(* Logix 5000 project; controller CIP vendor 1 type 14 code 106 rev 20.12; software revision 20.06 *)

TASK MainTask (continuous, watchdog 500 ms) : MainProgram

MODULES
   Local : vendor 1 type 14 code 106 (Compact 0, rev 20.12)
      Digital_Input_2 : 1769-IQ16 (Compact 5, rev 3.1, Input RPI 20 ms)
      Digital_Input_3 : 1769-IQ16 (Compact 6, rev 3.1, Input RPI 20 ms)
      Digital_Input_1 : 1769-IQ16 (Compact 4, rev 3.1, Input RPI 20 ms)
      Analog_Output_1 : vendor 1 type 10 code 45 (Compact 3, rev 2.1, Output RPI 80 ms)
      Analog_Input_1 : 1769-IF8 (Compact 1, rev 1.1, Output RPI 80 ms)
      Digital_Output_2 : 1769-OB16 (Compact 8, rev 3.1, Output RPI 20 ms)
      Analog_Input_2 : 1769-IF8 (Compact 2, rev 1.1, Output RPI 80 ms)
      Digital_Output_1 : 1769-OB16 (Compact 7, rev 3.1, Output RPI 20 ms)
      WASHER : 1734-AENT (Ethernet 192.168.1.58, rev 4.3, Output RPI 20 ms)
         Washer_Digital_Input_3 : 1734-IB8 (PointIO 5, rev 3.22)
         Washer_Digital_Input_1 : 1734-IB8 (PointIO 3, rev 3.22)
         Washer_Digital_Input_2 : 1734-IB8 (PointIO 4, rev 3.22)
         Washer_Analog_Input_1 : vendor 1 type 115 code 210 (PointIO 1, rev 3.2, Input RPI 80 ms)
         Washer_Digital_Output_2 : 1734-OB8 (PointIO 7, rev 3.22)
         Washer_Analog_Output_1 : 1734-OE2C (PointIO 2, rev 3.5, Output RPI 80 ms)
         Washer_Digital_Output_3 : 1734-OB8 (PointIO 8, rev 3.22)
         Washer_Digital_Output_1 : 1734-OB8 (PointIO 6, rev 3.22)
END_MODULES

TYPE Produce_Consume_Data :
STRUCT
   CommStatus : CONNECTION_STATUS;
   String : STRING[2];
   Real : REAL[10];
   DINT : DINT[10];
END_STRUCT
END_TYPE

TYPE RECIPE :
STRUCT
   OpCode : DINT[97];
   StepTime : DINT[97];
   Setpoint : REAL[97];
   Name : STRING;
END_STRUCT
END_TYPE

TYPE Security_Main_HMI :
STRUCT
   Timers : TIMER[10];
   Bits : DINT;
   Counters : COUNTER[6];
   User_Security_Name : STRING;
   User_Security_Name_Display : STRING[2];
   User_Security_Name_Temp : STRING;
   User_Security_Password : STRING;
   User_Security_Password_Temp : STRING;
   User_Security_Level : DINT;
   Number_Of_Users : DINT;
   User_Names : STRING[53];
   User_Names_Edit : STRING[53];
   User_Passwords : STRING[53];
   User_Passwords_Edit : STRING[53];
   User_Security_Levels : DINT[53];
   User_Security_Levels_Edit : DINT[53];
   Security_Save_Edit_Changes : BOOL;
   Security_Login_Enter_User_Button : BOOL;
   Security_Logout_Button : BOOL;
   Control_1 : CONTROL;
   Control_2 : CONTROL;
   Control_3 : CONTROL;
   User_Security_Name_Clear : STRING;
   User_Security_Password_Clear : STRING;
   Security_Login_Enter_Password_Button : BOOL;
   Name_Temp : DINT;
   Password_Temp : DINT;
   Auto_Logout_Counter : COUNTER;
   Auto_Logout_Timer_Enable : BOOL;
   Auto_Logout_Timer_Enabled : BOOL;
   Auto_Logout_Preset : DINT;
   Auto_Logout_Temp : DINT;
   PanelView_Control : DINT;
   PanelView_Status : DINT;
   PanelView_Security_Edit_Active : BOOL;
   PanelView_Security_Password_Length : DINT;
END_STRUCT
END_TYPE

TYPE Security_Remote_HMI :
STRUCT
   Timers : TIMER[3];
   Bits : DINT;
   User_Security_Name : STRING;
   User_Security_Name_Display : STRING[2];
   User_Security_Name_Temp : STRING;
   User_Security_Password : STRING;
   User_Security_Password_Temp : STRING;
   User_Security_Level : DINT;
   Number_Of_Users : DINT;
   User_Names : STRING[53];
   User_Passwords : STRING[53];
   User_Security_Levels : DINT[53];
   Security_Login_Enter_User_Button : BOOL;
   Security_Logout_Button : BOOL;
   Control_1 : CONTROL;
   User_Security_Name_Clear : STRING;
   User_Security_Password_Clear : STRING;
   Security_Login_Enter_Password_Button : BOOL;
   Auto_Logout_Counter : COUNTER;
   Auto_Logout_Timer_Enable : BOOL;
   Auto_Logout_Timer_Enabled : BOOL;
   Auto_Logout_Temp : DINT;
   PanelView_Control : DINT;
   PanelView_Status : DINT;
END_STRUCT
END_TYPE

VAR_GLOBAL   (* controller tags *)
   Alarm_Ack : INT[8];
   Alarm_Ack_All_PB : BOOL;
   Alarm_Present : INT[8] := ([0] := 70, [7] := 16384);
   Alarm_Preset_Indx : DINT := 118;
   Alarm_Remote_Ack_All : BOOL;
   Alarm_Status_Reset : BOOL;
   Alarm_Timer : TIMER[128] := ([0].PRE := 1500, [1].ACC := 4, [1].EN := 1, [1].DN := 1, [2].ACC := 4, [2].EN := 1, [2].DN := 1, [6].PRE := 3000, [7].PRE := 5000, [8].PRE := 5000, [9].PRE := 5000, [10].PRE := 5000, [11].PRE := 5000, [12].PRE := 5000, [13].PRE := 5000, [14].PRE := 5000, [15].PRE := 5000, [16].PRE := 5000, [17].PRE := 5000, [17].ACC := 5000, [17].EN := 1, [17].DN := 1, [18].PRE := 3000000, [19].PRE := 300000, [20].PRE := 1000, [21].PRE := 5000, [22].PRE := 1000, [23].PRE := 300000, [24].PRE := 900000, [25].PRE := 900000, [26].PRE := 300000, [27].PRE := 300000, [28].PRE := 500, [29].PRE := 500, [30].PRE := 8000, [31].PRE := 15000, [32].PRE := 8000, [33].PRE := 15000, [34].PRE := 8000, [35].PRE := 15000, [36].PRE := 8000, [37].PRE := 15000, [38].PRE := 5000, [39].PRE := 5000, [40].PRE := 3000, [41].PRE := 3000, [42].PRE := 3000, [44].PRE := 300000, [45].PRE := 5000, [45].ACC := 5001, [45].EN := 1, [45].DN := 1, [46].PRE := 8000, [47].PRE := 15000, [48].PRE := 8000, [49].PRE := 15000, [50].PRE := 5000, [51].PRE := 5000, [52].PRE := 5000, [53].PRE := 5000,
        [54].PRE := 5000, [55].PRE := 5000, [56].PRE := 5000, [57].PRE := 5000, [58].PRE := 5000, [59].PRE := 5000, [60].PRE := 5000, [61].PRE := 5000, [62].PRE := 5000, [63].PRE := 5000, [64].PRE := 5000, [65].PRE := 5000, [66].PRE := 5000, [67].PRE := 5000, [68].PRE := 5000, [69].PRE := 5000, [70].PRE := 5000, [71].PRE := 5000, [72].PRE := 5000, [73].PRE := 5000, [74].PRE := 5000, [75].PRE := 5000, [76].PRE := 5000, [77].PRE := 5000, [78].PRE := 5000, [78].ACC := 5001, [78].EN := 1, [78].DN := 1, [79].PRE := 5000, [79].ACC := 5001, [79].EN := 1, [79].DN := 1, [80].PRE := 5000, [81].PRE := 5000, [82].PRE := 5000, [83].PRE := 5000, [83].ACC := 5001, [83].EN := 1, [83].DN := 1, [84].PRE := 3000, [85].PRE := 3000, [85].ACC := 3002, [85].EN := 1, [85].DN := 1, [86].PRE := 1000, [87].PRE := 3000, [88].PRE := 10000, [89].PRE := 1800000, [90].PRE := 3000, [91].PRE := 3000, [93].PRE := 20000, [94].PRE := 10000, [95].PRE := 1000, [96].PRE := 5000, [96].ACC := 5001, [96].EN := 1, [96].DN := 1, [97].PRE := 5000, [97].ACC := 5001, [97].EN := 1,
        [97].DN := 1, [98].PRE := 5000, [98].ACC := 5001, [98].EN := 1, [98].DN := 1, [99].PRE := 5000, [99].ACC := 5001, [99].EN := 1, [99].DN := 1, [100].PRE := 10000, [101].PRE := 10000, [102].PRE := 10000, [103].PRE := 10000, [104].PRE := 5000, [105].PRE := 5000, [106].PRE := 5000, [107].PRE := 5000, [108].PRE := 5000, [109].PRE := 5000, [110].PRE := 5000, [111].PRE := 5000, [112].PRE := 5000, [113].PRE := 5000, [114].PRE := 5000, [114].ACC := 5001, [114].EN := 1, [114].DN := 1, [115].PRE := 5000, [115].ACC := 5001, [115].EN := 1, [115].DN := 1, [116].PRE := 8000, [117].PRE := 15000, [118].PRE := 8000, [119].PRE := 15000, [120].PRE := 8000, [121].PRE := 15000, [122].PRE := 8000, [123].PRE := 15000, [124].PRE := 5000, [124].ACC := 5001, [124].EN := 1, [124].DN := 1, [125].PRE := 5000, [125].ACC := 5001, [125].EN := 1, [125].DN := 1, [126].PRE := 5000, [126].ACC := 576, [126].EN := 1, [126].TT := 1, [127].PRE := 5000, [127].ACC := 5001, [127].EN := 1, [127].DN := 1);
   Alarm_Timer_Preset : DINT[128] := ([6] := 3000, [7] := 5000, [8] := 5000, [9] := 5000, [10] := 5000, [11] := 5000, [12] := 5000, [13] := 5000, [14] := 5000, [15] := 5000, [16] := 5000, [17] := 5000, [18] := 3000000, [19] := 300000, [20] := 1000, [21] := 5000, [22] := 1000, [23] := 300000, [24] := 900000, [25] := 900000, [26] := 300000, [27] := 300000, [28] := 500, [29] := 500, [30] := 8000, [31] := 15000, [32] := 8000, [33] := 15000, [34] := 8000, [35] := 15000, [36] := 8000, [37] := 15000, [38] := 5000, [39] := 5000, [40] := 3000, [41] := 3000, [42] := 3000, [44] := 300000, [45] := 5000, [46] := 8000, [47] := 15000, [48] := 8000, [49] := 15000, [50] := 5000, [51] := 5000, [52] := 5000, [53] := 5000, [54] := 5000, [55] := 5000, [56] := 5000, [57] := 5000, [58] := 5000, [59] := 5000, [60] := 5000, [61] := 5000, [62] := 5000, [63] := 5000, [64] := 5000, [65] := 5000, [66] := 5000,
        [67] := 5000, [68] := 5000, [69] := 5000, [70] := 5000, [71] := 5000, [72] := 5000, [73] := 5000, [74] := 5000, [75] := 5000, [76] := 5000, [77] := 5000, [78] := 5000, [79] := 5000, [80] := 5000, [81] := 5000, [82] := 5000, [83] := 5000, [84] := 3000, [85] := 3000, [86] := 1000, [87] := 3000, [88] := 10000, [89] := 1800000, [90] := 3000, [91] := 3000, [93] := 20000, [94] := 10000, [95] := 1000, [96] := 5000, [97] := 5000, [98] := 5000, [99] := 5000, [100] := 10000, [101] := 10000, [102] := 10000, [103] := 10000, [104] := 5000, [105] := 5000, [106] := 5000, [107] := 5000, [108] := 5000, [109] := 5000, [110] := 5000, [111] := 5000, [112] := 5000, [113] := 5000, [114] := 5000, [115] := 5000, [116] := 8000, [117] := 15000, [118] := 8000, [119] := 15000, [120] := 8000, [121] := 15000, [122] := 8000, [123] := 15000, [124] := 5000, [125] := 5000, [126] := 5000, [127] := 5000);
   Bit : BOOL[128] := ([10] := 1, [15] := 1, [16] := 1, [30] := 1, [34] := 1, [35] := 1, [37] := 1, [40] := 1, [41] := 1, [49] := 1, [52] := 1, [54] := 1, [55] := 1, [60] := 1, [66] := 1, [68] := 1, [70] := 1, [81] := 1, [82] := 1, [100] := 1);
   Counter : COUNTER[10] := ([1].PRE := 9999, [1].ACC := 1, [2].PRE := 4, [3].PRE := 3, [5].PRE := 64, [5].ACC := 12, [6].PRE := 20);
   IN_F8_50_99 : REAL[50] := ([0] := nan); {produced}
   IN_N7_100_199 : INT[100] := ([0] := 35, [1] := 1, [50] := 22428, [51] := -3734, [52] := 32, [53] := -32768, [54] := 12, [55] := -32768, [56] := 11180, [57] := -3792, [58] := 4804, [59] := 976, [60] := 16578, [61] := 20792, [62] := 1, [64] := 4, [66] := 3, [74] := 1, [76] := 12, [77] := -32768, [78] := 12, [79] := -32768, [80] := 11180, [81] := -3792, [82] := 30396, [83] := 1, [84] := 16578, [85] := 19059, [86] := 1, [88] := 4, [90] := 3); {produced}
   Integer : DINT[150] := ([0] := 1, [1] := 1, [5] := 2, [6] := 2, [7] := 1, [8] := 7, [10] := 36, [11] := 29, [12] := 65, [15] := -33, [20] := 20, [21] := 21, [22] := 61, [26] := 120, [27] := 120, [28] := 100, [29] := 1, [36] := -4, [38] := -1, [39] := 190, [40] := 80, [41] := 80, [43] := 120, [44] := 120, [45] := 120, [46] := 120, [48] := 50, [52] := 2, [53] := -2, [54] := 2, [56] := 6242, [57] := 31208, [58] := 12, [60] := 16383, [61] := 84, [62] := 10000, [80] := 5921);
   Integer_1 : ALIAS FOR Integer[1];
   Integer_6 : ALIAS FOR Integer[6];
   IO_Status : INT := 16384;
   IO_Status_Masked : INT := 16384;
   Level_Bits : BOOL[32] := ([1] := 1, [3] := 1, [4] := 1, [5] := 1, [7] := 1, [10] := 1, [11] := 1, [15] := 1, [17] := 1, [18] := 1, [19] := 1, [20] := 1);
   Level_Timers : TIMER[20] := ([0].PRE := 30000, [1].PRE := 60000, [2].PRE := 45000, [3].PRE := 75000, [3].ACC := 3, [3].EN := 1, [3].DN := 1, [4].PRE := 900000, [4].ACC := 900004, [4].EN := 1, [4].DN := 1, [5].PRE := 75000, [5].ACC := 75001, [5].EN := 1, [5].DN := 1, [7].PRE := 3000, [7].ACC := 3002, [7].EN := 1, [7].DN := 1, [8].PRE := 3000, [8].ACC := 3000, [8].EN := 1, [8].DN := 1, [10].PRE := 2000, [11].PRE := 1000, [11].ACC := 1000, [12].PRE := 1000, [12].ACC := 1000, [13].PRE := 1000, [13].ACC := 1000, [14].PRE := 1000, [14].ACC := 1000);
   Message_Index : ALIAS FOR Integer[30];
   Message_Present : INT[4] := ([1] := -32768, [3] := 2048);
   Message_SEQ : DINT[101] := ([1] := 32, [2] := 32, [3] := 14, [4] := 31, [5] := 32, [6] := 25, [7] := 36);
   Message_Timer : TIMER[1] := ([0].PRE := 1500, [0].ACC := 89, [0].EN := 1, [0].TT := 1);
   Minor_Faults : DINT;
   MOA_OFF : DINT[10] := ([1] := 2112);
   MOA_ON : DINT[10] := ([1] := 8320, [2] := 1536);
   MOA_ONS : DINT;
   MOA_Screen1_Auto : BOOL;
   MOA_Screen1_Man_Off : BOOL;
   MOA_Screen1_Man_On : BOOL;
   MOA_Screen2_Auto : BOOL;
   MOA_Screen2_Man_Off : BOOL;
   MOA_Screen2_Man_On : BOOL;
   MOA_Screen3_Auto : BOOL;
   MOA_Screen3_Man_Off : BOOL;
   MOA_Screen3_Man_On : BOOL;
   MOA_Screen4_Auto : BOOL;
   MOA_Screen4_Man_Off : BOOL;
   MOA_Screen4_Man_On : BOOL;
   MOA_Select : DINT[10] := ([1] := 8192, [2] := 1024, [3] := 64, [4] := 128, [5] := 128, [6] := 1);
   MOA_SP_Supply_Pump_Speed : DINT := 35;
   MOA_Status : DINT[10] := ([1] := 10432, [2] := 1536);
   MOA_Temp : DINT := -1025;
   One_Shot : BOOL[128] := ([11] := 1, [12] := 1, [13] := 1, [14] := 1, [15] := 1, [16] := 1, [17] := 1, [29] := 1, [30] := 1, [31] := 1, [32] := 1, [50] := 1);
   OpCode_Pin : DINT[5];
   OpCode_Word : DINT[5,97] := ([1,2] := 16#0000_821c, [1,3] := 16#0000_823c, [1,4] := 16#0000_823c, [1,5] := 16#0000_2001, [1,6] := 16#0000_0004, [1,8] := 16#0000_803d, [1,9] := 16#0000_0125, [1,10] := 16#0000_0125, [1,11] := 16#0000_0125, [1,12] := 16#0000_0125, [1,13] := 16#0000_180c, [1,14] := 16#0000_180c, [1,15] := 16#0000_180c, [1,16] := 16#0000_180c, [1,17] := 16#0000_180c, [1,18] := 16#0000_180c, [1,19] := 16#0000_180c, [1,20] := 16#0000_180c, [1,21] := 16#0000_0025, [1,22] := 16#0000_0025, [1,23] := 16#0000_0025, [1,24] := 16#0000_0025, [1,25] := 16#0000_100c, [1,26] := 16#0000_100c, [1,27] := 16#0000_100c, [1,28] := 16#0000_100c, [1,29] := 16#0000_0525, [1,30] := 16#0000_0525, [1,31] := 16#0000_0525, [1,32] := 16#0000_0525, [1,33] := 16#0000_1804, [1,34] := 16#0000_1804, [1,37] := 16#0000_8224, [1,38] := 16#0000_8224, [1,39] := 16#0000_8224, [1,40] := 16#0000_8020, [1,41] := 16#0000_8020, [1,42] := 16#0000_8020, [1,43] := 16#0000_80a0, [1,44] := 16#0000_80a0, [1,45] := 16#0000_80a0, [1,46] := 16#0000_8080, [1,47] := 16#0000_8080, [1,55] := 16#0000_0005, [1,56] := 16#0000_8204, [1,57] := 16#0000_8204, [1,58] := 16#0000_0005, [1,59] := 16#0000_0005, [1,60] := 16#0000_8080, [2,6] := 16#0000_8000, [2,9] := 16#0000_c800, [2,10] := 16#0000_c800, [2,11] := 16#0000_c800, [2,12] := 16#0000_c800, [2,13] := 16#0000_c202, [2,14] := 16#0000_c202, [2,15] := 16#0000_c202, [2,16] := 16#0000_c202, [2,17] := 16#0000_c101, [2,18] := 16#0000_c101,
        [2,19] := 16#0000_c101, [2,20] := 16#0000_c101, [2,21] := 16#0000_c400, [2,22] := 16#0000_c400, [2,23] := 16#0000_c400, [2,24] := 16#0000_c400, [2,25] := 16#0000_c400, [2,26] := 16#0000_c400, [2,27] := 16#0000_c400, [2,28] := 16#0000_c400, [2,29] := 16#0000_c080, [2,30] := 16#0000_c080, [2,31] := 16#0000_c080, [2,32] := 16#0000_c080, [2,33] := 16#0000_8202, [2,34] := 16#0000_8101, [2,37] := 16#0000_c000, [2,38] := 16#0000_c000, [2,39] := 16#0000_c000, [2,40] := 16#0000_4000, [2,41] := 16#0000_4000, [2,42] := 16#0000_4000, [2,43] := 16#0000_4000, [2,44] := 16#0000_4000, [2,45] := 16#0000_4000, [2,55] := 16#0000_8800, [2,56] := 16#0000_8200, [2,57] := 16#0000_8100, [2,58] := 16#0000_8400, [2,59] := 16#0000_8080, [3,2] := 16#0000_4020, [3,3] := 16#0000_f2f0, [3,4] := 16#0000_cd30, [3,5] := 16#0000_4000, [3,6] := 16#0000_4000, [3,8] := 16#0000_0020, [3,9] := 16#0000_a200, [3,10] := 16#0000_9200, [3,11] := 16#0000_8900, [3,12] := 16#0000_8500, [3,13] := 16#0000_a200, [3,14] := 16#0000_9200, [3,15] := 16#0000_8900, [3,16] := 16#0000_8500, [3,17] := 16#0000_a200, [3,18] := 16#0000_9200, [3,19] := 16#0000_8900, [3,20] := 16#0000_8500, [3,21] := 16#0000_a200, [3,22] := 16#0000_9200, [3,23] := 16#0000_8900, [3,24] := 16#0000_8500, [3,25] := 16#0000_a200, [3,26] := 16#0000_9200, [3,27] := 16#0000_8900, [3,28] := 16#0000_8500, [3,29] := 16#0000_a200, [3,30] := 16#0000_9200, [3,31] := 16#0000_8900, [3,32] := 16#0000_8500,
        [3,33] := 16#0000_4000, [3,34] := 16#0000_4000, [3,35] := 16#0000_3210, [3,36] := 16#0000_3210, [3,37] := 16#0000_b200, [3,38] := 16#0000_8900, [3,39] := 16#0000_8500, [3,40] := 16#0000_0200, [3,41] := 16#0000_0100, [3,42] := 16#0000_0100, [3,43] := 16#0000_3200, [3,44] := 16#0000_0900, [3,45] := 16#0000_0500, [3,46] := 16#0000_2080, [3,47] := 16#0000_1040, [3,55] := 16#0000_8008, [3,56] := 16#0000_8008, [3,57] := 16#0000_8008, [3,58] := 16#0000_8008, [3,59] := 16#0000_8008, [3,60] := 16#0000_0008, [3,65] := 16#0000_0001, [3,66] := 16#0000_0001, [3,67] := 16#0000_0001, [3,68] := 16#0000_0001, [3,69] := 16#0000_0001, [4,35] := 16#0000_0003, [4,36] := 16#0000_0001, [4,49] := 16#0000_2000, [4,50] := 16#0000_1000, [4,51] := 16#0000_0800, [4,52] := 16#0000_0400, [4,53] := 16#0000_0200, [4,54] := 16#0000_0100);
   OUT_F8_0_49 : REAL[50] := ([1] := 21.79088, [2] := 22.761398, [5] := 14.0, [6] := 3.1312947, [7] := -0.5218824, [8] := -1.4997253, [9] := 0.003662333, [11] := 20.120556, [12] := 20.04044, [20] := 50.0, [30] := 60.0, [31] := 0.2, [32] := 0.1, [33] := 110.0, [34] := 195.0, [35] := 10.0, [36] := 150.0, [37] := 190.0, [38] := 60.0, [39] := 60.0, [40] := 80.0, [41] := 190.0, [42] := 5.5, [43] := 10.5); {produced}
   OUT_N7_0_99 : INT[100] := ([0] := 4, [1] := 8, [2] := 1, [6] := 32, [10] := 12, [11] := -21846, [12] := 2730, [13] := 8320, [14] := 1536, [20] := 20482, [21] := 170, [22] := 8, [30] := 70, [37] := 16384, [41] := -32768); {produced}
   Panelview : INT[40] := ([0] := 6144, [3] := 65, [8] := 1, [14] := 1, [15] := 1, [20] := 2, [31] := 1, [32] := 1, [33] := 1, [34] := -1);
   PID1 : PID := (CTL := -2080340864, EN := 1, SWM := 1, INI := 1, DVNA := 1, PVHA := 1, KP := 1.2, KI := 0.1, BIAS := 46.65812, MAXS := 100.0, MAXO := 51.0, UPD := 0.01, PV := 21.79088, ERR := -21.79088, MAXI := 100.0, MAXCV := 16383.0, MAXTIE := 16383.0, DATA[0] := -20.509062, DATA[1] := -348.65408, DATA[2] := 21.79088, DATA[3] := -21.79088, DATA[5] := 1.0, DATA[6] := 1.0, DATA[7] := 0.16, DATA[8] := 1.2, DATA[9] := 0.1, DATA[11] := 1.2, DATA[12] := 0.1, DATA[15] := 163.83, DATA[16] := 0.006103888);
   PID2 : PID := (CTL := -2080340864, EN := 1, SWM := 1, INI := 1, DVNA := 1, PVHA := 1, KP := 0.5, KI := 0.125, BIAS := 1.0468168, MAXS := 150.0, MAXO := 100.0, UPD := 0.01, PV := 3.1312947, ERR := -3.1312947, MAXI := 150.0, MAXCV := 16383.0, MAXTIE := 16383.0, DATA[0] := -0.003051877, DATA[1] := -33.40048, DATA[2] := 3.1312947, DATA[3] := -3.1312947, DATA[5] := 0.6666667, DATA[6] := 1.0, DATA[7] := 0.16, DATA[8] := 0.5, DATA[9] := 0.125, DATA[11] := 0.5, DATA[12] := 0.125, DATA[15] := 163.83, DATA[16] := 0.006103888);
   PID3 : PID := (CTL := -2080340864, EN := 1, SWM := 1, INI := 1, DVNA := 1, PVHA := 1, KP := 8.0, KI := 0.1, BIAS := 75.446365, MAXS := 150.0, DB := 3.0, MAXO := 100.0, UPD := 0.01, PV := 20.120556, ERR := -20.120556, MAXI := 150.0, MAXCV := 16383.0, MAXTIE := 16383.0, DATA[0] := 31.863266, DATA[1] := -214.61926, DATA[2] := 20.120556, DATA[3] := -20.120556, DATA[5] := 0.6666667, DATA[6] := 1.0, DATA[7] := 0.16, DATA[8] := 8.0, DATA[9] := 0.1, DATA[11] := 8.0, DATA[12] := 0.1, DATA[15] := 163.83, DATA[16] := 0.006103888);
   PID3_Timer : TIMER[4] := ([0].PRE := 5000);
   PID_Button : DINT[5];
   PID_Button_ONS : DINT[5];
   PID_ONS : DINT[5] := ([1] := 2, [2] := 10, [3] := 2, [4] := 4);
   PID_Timer : TIMER[5] := ([0].PRE := 5000, [0].ACC := 5000, [0].EN := 1, [0].DN := 1, [1].PRE := 10000, [2].PRE := 5000, [2].EN := 1, [2].DN := 1, [3].PRE := 4000, [4].PRE := 50, [4].ACC := 53, [4].EN := 1, [4].DN := 1);
   PV_Current_Select_Step_Op : DINT := 52;
   PV_Edit_Opcodes : DINT[300] := ([1] := 50, [2] := 5, [3] := 52, [4] := 12, [5] := 11, [6] := 65, [7] := 41, [8] := 5, [9] := 33, [10] := 16, [11] := 15, [12] := 67, [13] := 38, [14] := 41, [15] := 2, [16] := 8, [17] := 51, [18] := 5, [19] := 6, [20] := 28, [21] := 27, [22] := 66, [23] := 38, [24] := 41, [25] := 2, [26] := 8, [27] := 49, [28] := 5, [29] := 24, [30] := 23, [31] := 66, [32] := 5, [33] := 32, [34] := 31, [35] := 69, [36] := 2, [37] := 44, [38] := 45, [39] := 4, [40] := 1, [101] := 10, [201] := 24, [202] := 66, [203] := 49, [204] := 5, [205] := 32, [206] := 69, [207] := 45, [208] := 2, [209] := 1, [287] := 10);
   PV_Edit_Recipe_Name : STRING := 'TANK WASH W/DIP TUBES CYCLE #2';
   PV_Edit_Recipe_Top_Row : DINT := 1;
   PV_Edit_Recipes : DINT[7] := ([0] := 3, [1] := 52, [2] := 1, [4] := 1);
   PV_Edit_Recipes_0 : ALIAS FOR PV_Edit_Recipes[0];
   PV_Edit_Recipes_0_Prev : DINT;
   PV_Edit_Screen_Opcodes : DINT[17] := ([1] := 50, [2] := 5, [3] := 52, [4] := 12, [5] := 11, [6] := 65, [7] := 41, [8] := 5, [9] := 33, [10] := 16, [11] := 15, [12] := 67, [13] := 38, [14] := 41, [15] := 2, [16] := 8);
   PV_Edit_Setpoints : REAL[97] := ([1] := 45.0, [2] := 45.0, [3] := 45.0, [4] := 45.0, [5] := 45.0, [6] := 25.0, [7] := 42.0, [8] := 42.0, [9] := 42.0, [10] := 42.0, [11] := 42.0, [12] := 22.0, [13] := 60.0, [14] := 900.0, [15] := 300.0, [16] := 300.0, [17] := 5.0, [18] := 4.5, [19] := 30.0, [20] := 60.0, [21] := 5.0, [22] := 15.0, [23] := 300.0, [24] := 0.2, [25] := 2.0, [26] := 1.5, [27] := 60.0, [28] := 50.0, [29] := 30.0, [30] := 30.0, [31] := 300.0, [32] := 0.1, [33] := 5.0, [34] := 900.0, [37] := 70.0, [38] := 100.0, [39] := 110.0, [40] := 30.0, [41] := 60.0, [42] := 900.0, [43] := 3000.0, [44] := 300.0, [45] := 195.0, [46] := 10.0, [47] := 150.0, [48] := 190.0, [49] := 60.0, [50] := 60.0, [51] := 80.0, [52] := 190.0, [53] := 50.0, [54] := 85.0, [55] := 40.0, [56] := 25.0, [57] := 10.0, [58] := 4.0, [61] := 5.0, [62] := 1.0, [65] := 100.0, [66] := 15.0,
        [67] := 50.0, [68] := 5.0, [69] := 60.0, [70] := 20.0, [71] := 60.0, [72] := 2.0, [73] := 120.0, [74] := 20.0, [75] := 120.0, [76] := 20.0, [77] := 40.0, [78] := 15.0, [79] := 30.0, [80] := 5.0, [81] := 45.0, [82] := 30.0, [83] := 5.0, [85] := 5.5, [86] := 10.5, [92] := 75.0, [93] := 90.0, [94] := 5.0, [95] := 110.0, [96] := 10.0);
   PV_Edit_Times : DINT[300] := ([1] := 1, [2] := 1, [3] := 1, [4] := 10, [5] := 70, [6] := 1, [7] := 3, [8] := 1, [9] := 30, [10] := 50, [11] := 150, [12] := 1, [13] := 3, [14] := 3, [15] := 10, [16] := 20, [17] := 1, [18] := 1, [19] := 3, [20] := 15, [21] := 50, [22] := 1, [23] := 1, [24] := 3, [25] := 10, [26] := 20, [27] := 1, [28] := 1, [29] := 20, [30] := 40, [31] := 1, [32] := 1, [33] := 10, [34] := 10, [35] := 1, [36] := 10, [37] := 20, [38] := 20, [39] := 10, [40] := 1, [201] := 20, [202] := 1, [203] := 1, [204] := 1, [205] := 10, [206] := 1, [207] := 10, [208] := 10, [209] := 1);
   PV_Message : DINT[3] := ([0] := 32, [2] := 5);
   PV_Output_Status : INT[10] := ([1] := 8320, [2] := 1536, [3] := 8);
   PV_Output_Status_IND : INT[10,16] := ([1,7] := 1, [1,13] := 1, [2,9] := 1, [2,10] := 1, [3,3] := 1);
   PV_Rename_Recipe_Name : STRING := 'TANK WASH W/DIP TUBES CYCLE #2';
   PV_Security : Security_Main_HMI := (Timers[0].PRE := 2000, Timers[1].PRE := 2000, Timers[2].PRE := 25, Timers[2].ACC := 4, Timers[2].EN := 1, Timers[2].TT := 1, Timers[3].PRE := 3000, Timers[3].ACC := 3001, Timers[3].EN := 1, Timers[3].DN := 1, Timers[4].PRE := 25, Timers[4].ACC := 25, Timers[4].EN := 1, Timers[4].DN := 1, Timers[5].PRE := 2000, Timers[5].ACC := 2002, Timers[5].EN := 1, Timers[5].DN := 1, Timers[6].PRE := 60000, Timers[7].PRE := 2000, Timers[8].PRE := 3000, Timers[9].PRE := 200, Bits := 1179648, Counters[0].PRE := 9999, Counters[0].ACC := 1, Counters[0].CU := 1, Counters[1].PRE := 53, Counters[1].ACC := 48, Counters[2].PRE := 9999, Counters[3].PRE := 53, Counters[3].ACC := 5, Counters[3].CU := 1, User_Security_Name := 'DEFAULT', User_Security_Name_Display[0] := 'DEFAULT', User_Security_Password_Temp := '1', Number_Of_Users := 52, User_Names[1] := '1', User_Names[2] := '2', User_Names[3] := '3', User_Names[4] := '4', User_Names[5] := '5', User_Names[6] := '6', User_Names[7] := '7', User_Names[8] := '8', User_Names[9] := '9', User_Names[10] := '10', User_Names[11] := '11', User_Names[12] := '12', User_Names[13] := '13', User_Names[14] := '14', User_Names[15] := '15', User_Names[16] := '16', User_Names[17] := '17', User_Names[18] := '18', User_Names[19] := '19', User_Names[20] := '20', User_Names[21] := '21', User_Names[22] := '22', User_Names[23] := '23', User_Names[24] := '24',
        User_Names[25] := '25', User_Names[26] := '26', User_Names[27] := '27', User_Names[28] := '28', User_Names[29] := '29', User_Names[30] := '30', User_Names[31] := '31', User_Names[32] := '32', User_Names[33] := '33', User_Names[34] := '34', User_Names[35] := '35', User_Names[36] := '36', User_Names[37] := '37', User_Names[38] := '38', User_Names[39] := '39', User_Names[40] := '40', User_Names[41] := '41', User_Names[42] := '42', User_Names[43] := '43', User_Names[44] := '44', User_Names[45] := '45', User_Names[46] := '46', User_Names[47] := '47', User_Names[48] := '48', User_Names[49] := '49', User_Names[50] := '50', User_Names[51] := 'sanimatic', User_Names_Edit[1] := '1', User_Names_Edit[2] := '2', User_Names_Edit[3] := '3', User_Names_Edit[4] := '4', User_Names_Edit[5] := '5', User_Names_Edit[6] := '6', User_Names_Edit[7] := '7', User_Names_Edit[8] := '8', User_Names_Edit[9] := '9', User_Names_Edit[10] := '10', User_Names_Edit[11] := '11', User_Names_Edit[12] := '12', User_Names_Edit[13] := '13', User_Names_Edit[14] := '14', User_Names_Edit[15] := '15', User_Names_Edit[16] := '16', User_Names_Edit[17] := '17', User_Names_Edit[18] := '18', User_Names_Edit[19] := '19', User_Names_Edit[20] := '20', User_Names_Edit[21] := '21', User_Names_Edit[22] := '22', User_Names_Edit[23] := '23', User_Names_Edit[24] := '24', User_Names_Edit[25] := '25', User_Names_Edit[26] := '26', User_Names_Edit[27] := '27', User_Names_Edit[28] := '28', User_Names_Edit[29] := '29', User_Names_Edit[30] := '30', User_Names_Edit[31] := '31', User_Names_Edit[32] := '32', User_Names_Edit[33] := '33',
        User_Names_Edit[34] := '34', User_Names_Edit[35] := '35', User_Names_Edit[36] := '36', User_Names_Edit[37] := '37', User_Names_Edit[38] := '38', User_Names_Edit[39] := '39', User_Names_Edit[40] := '40', User_Names_Edit[41] := '41', User_Names_Edit[42] := '42', User_Names_Edit[43] := '43', User_Names_Edit[44] := '44', User_Names_Edit[45] := '45', User_Names_Edit[46] := '46', User_Names_Edit[47] := '47', User_Names_Edit[48] := '48', User_Names_Edit[49] := '49', User_Names_Edit[50] := '50', User_Names_Edit[51] := 'sanimatic', User_Passwords[1] := '1', User_Passwords[2] := '2', User_Passwords[3] := '3', User_Passwords[4] := '4', User_Passwords[5] := '5', User_Passwords[6] := '6', User_Passwords[7] := '7', User_Passwords[8] := '8', User_Passwords[9] := '9', User_Passwords[10] := '10', User_Passwords[11] := '11', User_Passwords[12] := '12', User_Passwords[13] := '13', User_Passwords[14] := '14', User_Passwords[15] := '15', User_Passwords[16] := '16', User_Passwords[17] := '17', User_Passwords[18] := '18', User_Passwords[19] := '19', User_Passwords[20] := '20', User_Passwords[21] := '21', User_Passwords[22] := '22', User_Passwords[23] := '23', User_Passwords[24] := '24', User_Passwords[25] := '25', User_Passwords[26] := '26', User_Passwords[27] := '27', User_Passwords[28] := '28', User_Passwords[29] := '29', User_Passwords[30] := '30', User_Passwords[31] := '31', User_Passwords[32] := '32', User_Passwords[33] := '33', User_Passwords[34] := '34', User_Passwords[35] := '35', User_Passwords[36] := '36', User_Passwords[37] := '37', User_Passwords[38] := '38', User_Passwords[39] := '39', User_Passwords[40] := '40', User_Passwords[41] := '41', User_Passwords[42] := '42',
        User_Passwords[43] := '43', User_Passwords[44] := '44', User_Passwords[45] := '45', User_Passwords[46] := '46', User_Passwords[47] := '47', User_Passwords[48] := '48', User_Passwords[49] := '49', User_Passwords[50] := '50', User_Passwords[51] := '1915', User_Passwords_Edit[1] := '1', User_Passwords_Edit[2] := '2', User_Passwords_Edit[3] := '3', User_Passwords_Edit[4] := '4', User_Passwords_Edit[5] := '5', User_Passwords_Edit[6] := '6', User_Passwords_Edit[7] := '7', User_Passwords_Edit[8] := '8', User_Passwords_Edit[9] := '9', User_Passwords_Edit[10] := '10', User_Passwords_Edit[11] := '11', User_Passwords_Edit[12] := '12', User_Passwords_Edit[13] := '13', User_Passwords_Edit[14] := '14', User_Passwords_Edit[15] := '15', User_Passwords_Edit[16] := '16', User_Passwords_Edit[17] := '17', User_Passwords_Edit[18] := '18', User_Passwords_Edit[19] := '19', User_Passwords_Edit[20] := '20', User_Passwords_Edit[21] := '21', User_Passwords_Edit[22] := '22', User_Passwords_Edit[23] := '23', User_Passwords_Edit[24] := '24', User_Passwords_Edit[25] := '25', User_Passwords_Edit[26] := '26', User_Passwords_Edit[27] := '27', User_Passwords_Edit[28] := '28', User_Passwords_Edit[29] := '29', User_Passwords_Edit[30] := '30', User_Passwords_Edit[31] := '31', User_Passwords_Edit[32] := '32', User_Passwords_Edit[33] := '33', User_Passwords_Edit[34] := '34', User_Passwords_Edit[35] := '35', User_Passwords_Edit[36] := '36', User_Passwords_Edit[37] := '37', User_Passwords_Edit[38] := '38', User_Passwords_Edit[39] := '39', User_Passwords_Edit[40] := '40', User_Passwords_Edit[41] := '41', User_Passwords_Edit[42] := '42', User_Passwords_Edit[43] := '43', User_Passwords_Edit[44] := '44', User_Passwords_Edit[45] := '45', User_Passwords_Edit[46] := '46', User_Passwords_Edit[47] := '47', User_Passwords_Edit[48] := '48', User_Passwords_Edit[49] := '49', User_Passwords_Edit[50] := '50', User_Passwords_Edit[51] := '1915',
        User_Security_Levels[1] := 1, User_Security_Levels[2] := 2, User_Security_Levels[3] := 3, User_Security_Levels[4] := 3, User_Security_Levels[47] := 3, User_Security_Levels[48] := 3, User_Security_Levels[49] := 3, User_Security_Levels[50] := 3, User_Security_Levels[51] := 3, User_Security_Levels_Edit[1] := 1, User_Security_Levels_Edit[2] := 2, User_Security_Levels_Edit[3] := 3, User_Security_Levels_Edit[4] := 3, User_Security_Levels_Edit[47] := 3, User_Security_Levels_Edit[48] := 3, User_Security_Levels_Edit[49] := 3, User_Security_Levels_Edit[50] := 3, User_Security_Levels_Edit[51] := 3, Control_1.LEN := 53, Control_1.POS := 52, Control_1.EN := 1, Control_1.DN := 1, Control_2.LEN := 53, Control_2.POS := 22, Control_2.EN := 1, Control_3.LEN := 53, Control_3.EN := 1, Control_3.IN := 1, Control_3.FD := 1, User_Security_Name_Clear := 'DEFAULT', Name_Temp := 3, Password_Temp := 36, Auto_Logout_Counter.PRE := 11, Auto_Logout_Preset := 11, Auto_Logout_Temp := 1, PanelView_Status := 1);
   PV_Security1 : Security_Remote_HMI := (Timers[0].PRE := 2000, Timers[1].PRE := 2000, Timers[2].PRE := 60000, Bits := 1196032, User_Security_Name := 'DEFAULT', User_Security_Name_Display[0] := 'DEFAULT', User_Security_Password_Temp := '4', Number_Of_Users := 52, User_Names[1] := '1', User_Names[2] := '2', User_Names[3] := '3', User_Names[4] := '4', User_Names[5] := '5', User_Names[6] := '6', User_Names[7] := '7', User_Names[8] := '8', User_Names[9] := '9', User_Names[10] := '10', User_Names[11] := '11', User_Names[12] := '12', User_Names[13] := '13', User_Names[14] := '14', User_Names[15] := '15', User_Names[16] := '16', User_Names[17] := '17', User_Names[18] := '18', User_Names[19] := '19', User_Names[20] := '20', User_Names[21] := '21', User_Names[22] := '22', User_Names[23] := '23', User_Names[24] := '24', User_Names[25] := '25', User_Names[26] := '26', User_Names[27] := '27', User_Names[28] := '28', User_Names[29] := '29', User_Names[30] := '30', User_Names[31] := '31', User_Names[32] := '32', User_Names[33] := '33', User_Names[34] := '34', User_Names[35] := '35', User_Names[36] := '36', User_Names[37] := '37', User_Names[38] := '38', User_Names[39] := '39', User_Names[40] := '40', User_Names[41] := '41', User_Names[42] := '42', User_Names[43] := '43', User_Names[44] := '44', User_Names[45] := '45', User_Names[46] := '46', User_Names[47] := '47', User_Names[48] := '48', User_Names[49] := '49', User_Names[50] := '50', User_Names[51] := 'sanimatic', User_Passwords[1] := '1',
        User_Passwords[2] := '2', User_Passwords[3] := '3', User_Passwords[4] := '4', User_Passwords[5] := '5', User_Passwords[6] := '6', User_Passwords[7] := '7', User_Passwords[8] := '8', User_Passwords[9] := '9', User_Passwords[10] := '10', User_Passwords[11] := '11', User_Passwords[12] := '12', User_Passwords[13] := '13', User_Passwords[14] := '14', User_Passwords[15] := '15', User_Passwords[16] := '16', User_Passwords[17] := '17', User_Passwords[18] := '18', User_Passwords[19] := '19', User_Passwords[20] := '20', User_Passwords[21] := '21', User_Passwords[22] := '22', User_Passwords[23] := '23', User_Passwords[24] := '24', User_Passwords[25] := '25', User_Passwords[26] := '26', User_Passwords[27] := '27', User_Passwords[28] := '28', User_Passwords[29] := '29', User_Passwords[30] := '30', User_Passwords[31] := '31', User_Passwords[32] := '32', User_Passwords[33] := '33', User_Passwords[34] := '34', User_Passwords[35] := '35', User_Passwords[36] := '36', User_Passwords[37] := '37', User_Passwords[38] := '38', User_Passwords[39] := '39', User_Passwords[40] := '40', User_Passwords[41] := '41', User_Passwords[42] := '42', User_Passwords[43] := '43', User_Passwords[44] := '44', User_Passwords[45] := '45', User_Passwords[46] := '46', User_Passwords[47] := '47', User_Passwords[48] := '48', User_Passwords[49] := '49', User_Passwords[50] := '50', User_Passwords[51] := '1915', User_Security_Levels[1] := 1, User_Security_Levels[2] := 2, User_Security_Levels[3] := 3, User_Security_Levels[4] := 3, User_Security_Levels[47] := 3, User_Security_Levels[48] := 3, User_Security_Levels[49] := 3, User_Security_Levels[50] := 3, User_Security_Levels[51] := 3, Control_1.LEN := 53,
        Control_1.POS := 13, Control_1.EN := 1, User_Security_Name_Clear := 'DEFAULT', Auto_Logout_Counter.PRE := 11, Auto_Logout_Timer_Enable := 1, Auto_Logout_Temp := 1, PanelView_Status := 1);
   PV_Status_Bit : BOOL := 1;
   PV_Step_Time : REAL;
   PV_Valve_Input_Status_IND : INT[10,16] := ([1,14] := 3, [1,15] := 3, [2,5] := 3, [2,6] := 3, [2,7] := 3, [2,8] := 3, [2,9] := 3, [2,10] := 3, [2,11] := 3, [2,12] := 3, [2,13] := 3, [2,14] := 3, [2,15] := 3);
   PV_Visibility : INT[5] := ([0] := 1069, [1] := 31, [3] := 3, [4] := 1205);
   PV_Visibility_Remote1_HMI : INT[5] := ([0] := 1069, [3] := 3);
   Recipe : RECIPE[41] := ([0].OpCode[1] := 50, [0].OpCode[2] := 5, [0].OpCode[3] := 52, [0].OpCode[4] := 12, [0].OpCode[5] := 11, [0].OpCode[6] := 65, [0].OpCode[7] := 41, [0].OpCode[8] := 5, [0].OpCode[9] := 33, [0].OpCode[10] := 16, [0].OpCode[11] := 15, [0].OpCode[12] := 67, [0].OpCode[13] := 38, [0].OpCode[14] := 41, [0].OpCode[15] := 2, [0].OpCode[16] := 8, [0].OpCode[17] := 51, [0].OpCode[18] := 5, [0].OpCode[19] := 6, [0].OpCode[20] := 28, [0].OpCode[21] := 27, [0].OpCode[22] := 66, [0].OpCode[23] := 38, [0].OpCode[24] := 41, [0].OpCode[25] := 2, [0].OpCode[26] := 8, [0].OpCode[27] := 49, [0].OpCode[28] := 5, [0].OpCode[29] := 24, [0].OpCode[30] := 23, [0].OpCode[31] := 66, [0].OpCode[32] := 5, [0].OpCode[33] := 32, [0].OpCode[34] := 31, [0].OpCode[35] := 69, [0].OpCode[36] := 2, [0].OpCode[37] := 44, [0].OpCode[38] := 45, [0].OpCode[39] := 4, [0].OpCode[40] := 1, [0].StepTime[1] := 1, [0].StepTime[2] := 1, [0].StepTime[3] := 1, [0].StepTime[4] := 10, [0].StepTime[5] := 70, [0].StepTime[6] := 1, [0].StepTime[7] := 3, [0].StepTime[8] := 1, [0].StepTime[9] := 30, [0].StepTime[10] := 50, [0].StepTime[11] := 150, [0].StepTime[12] := 1, [0].StepTime[13] := 3, [0].StepTime[14] := 3, [0].StepTime[15] := 10, [0].StepTime[16] := 20, [0].StepTime[17] := 1, [0].StepTime[18] := 1, [0].StepTime[19] := 3, [0].StepTime[20] := 15,
        [0].StepTime[21] := 50, [0].StepTime[22] := 1, [0].StepTime[23] := 1, [0].StepTime[24] := 3, [0].StepTime[25] := 10, [0].StepTime[26] := 20, [0].StepTime[27] := 1, [0].StepTime[28] := 1, [0].StepTime[29] := 20, [0].StepTime[30] := 40, [0].StepTime[31] := 1, [0].StepTime[32] := 1, [0].StepTime[33] := 10, [0].StepTime[34] := 10, [0].StepTime[35] := 1, [0].StepTime[36] := 10, [0].StepTime[37] := 20, [0].StepTime[38] := 20, [0].StepTime[39] := 10, [0].StepTime[40] := 1, [0].Setpoint[1] := 45.0, [0].Setpoint[2] := 45.0, [0].Setpoint[3] := 45.0, [0].Setpoint[4] := 45.0, [0].Setpoint[5] := 45.0, [0].Setpoint[6] := 25.0, [0].Setpoint[7] := 42.0, [0].Setpoint[8] := 42.0, [0].Setpoint[9] := 42.0, [0].Setpoint[10] := 42.0, [0].Setpoint[11] := 42.0, [0].Setpoint[12] := 22.0, [0].Setpoint[13] := 60.0, [0].Setpoint[14] := 900.0, [0].Setpoint[15] := 300.0, [0].Setpoint[16] := 300.0, [0].Setpoint[17] := 5.0, [0].Setpoint[18] := 4.5, [0].Setpoint[19] := 30.0, [0].Setpoint[20] := 60.0, [0].Setpoint[21] := 5.0, [0].Setpoint[22] := 15.0, [0].Setpoint[23] := 300.0, [0].Setpoint[24] := 0.2, [0].Setpoint[25] := 2.0, [0].Setpoint[26] := 1.5, [0].Setpoint[27] := 60.0, [0].Setpoint[28] := 50.0, [0].Setpoint[29] := 30.0, [0].Setpoint[30] := 30.0, [0].Setpoint[31] := 300.0, [0].Setpoint[32] := 0.1, [0].Setpoint[33] := 5.0, [0].Setpoint[34] := 900.0, [0].Setpoint[37] := 70.0, [0].Setpoint[38] := 100.0, [0].Setpoint[39] := 110.0, [0].Setpoint[40] := 30.0, [0].Setpoint[41] := 60.0, [0].Setpoint[42] := 900.0,
        [0].Setpoint[43] := 3000.0, [0].Setpoint[44] := 300.0, [0].Setpoint[45] := 195.0, [0].Setpoint[46] := 10.0, [0].Setpoint[47] := 150.0, [0].Setpoint[48] := 190.0, [0].Setpoint[49] := 60.0, [0].Setpoint[50] := 60.0, [0].Setpoint[51] := 80.0, [0].Setpoint[52] := 190.0, [0].Setpoint[53] := 50.0, [0].Setpoint[54] := 85.0, [0].Setpoint[55] := 40.0, [0].Setpoint[56] := 25.0, [0].Setpoint[57] := 10.0, [0].Setpoint[58] := 4.0, [0].Setpoint[61] := 5.0, [0].Setpoint[62] := 1.0, [0].Setpoint[65] := 100.0, [0].Setpoint[66] := 15.0, [0].Setpoint[67] := 50.0, [0].Setpoint[68] := 5.0, [0].Setpoint[69] := 60.0, [0].Setpoint[70] := 20.0, [0].Setpoint[71] := 60.0, [0].Setpoint[72] := 2.0, [0].Setpoint[73] := 120.0, [0].Setpoint[74] := 20.0, [0].Setpoint[75] := 120.0, [0].Setpoint[76] := 20.0, [0].Setpoint[77] := 40.0, [0].Setpoint[78] := 15.0, [0].Setpoint[79] := 30.0, [0].Setpoint[80] := 5.0, [0].Setpoint[81] := 45.0, [0].Setpoint[82] := 30.0, [0].Setpoint[83] := 5.0, [0].Setpoint[85] := 5.5, [0].Setpoint[86] := 10.5, [0].Setpoint[92] := 75.0, [0].Setpoint[93] := 90.0, [0].Setpoint[94] := 5.0, [0].Setpoint[95] := 110.0, [0].Setpoint[96] := 10.0, [0].Name := 'TANK WASH W/DIP TUBES CYCLE', [1].OpCode[1] := 50, [1].OpCode[2] := 5, [1].OpCode[3] := 52, [1].OpCode[4] := 12, [1].OpCode[5] := 11, [1].OpCode[6] := 65, [1].OpCode[7] := 41, [1].OpCode[8] := 5, [1].OpCode[9] := 33, [1].OpCode[10] := 16, [1].OpCode[11] := 15, [1].OpCode[12] := 67, [1].OpCode[13] := 38, [1].OpCode[14] := 41, [1].OpCode[15] := 2,
        [1].OpCode[16] := 8, [1].OpCode[17] := 51, [1].OpCode[18] := 5, [1].OpCode[19] := 6, [1].OpCode[20] := 28, [1].OpCode[21] := 27, [1].OpCode[22] := 66, [1].OpCode[23] := 38, [1].OpCode[24] := 41, [1].OpCode[25] := 2, [1].OpCode[26] := 8, [1].OpCode[27] := 49, [1].OpCode[28] := 5, [1].OpCode[29] := 24, [1].OpCode[30] := 23, [1].OpCode[31] := 66, [1].OpCode[32] := 5, [1].OpCode[33] := 32, [1].OpCode[34] := 31, [1].OpCode[35] := 69, [1].OpCode[36] := 2, [1].OpCode[37] := 44, [1].OpCode[38] := 45, [1].OpCode[39] := 4, [1].OpCode[40] := 1, [1].StepTime[1] := 1, [1].StepTime[2] := 1, [1].StepTime[3] := 1, [1].StepTime[4] := 10, [1].StepTime[5] := 70, [1].StepTime[6] := 1, [1].StepTime[7] := 3, [1].StepTime[8] := 1, [1].StepTime[9] := 30, [1].StepTime[10] := 50, [1].StepTime[11] := 150, [1].StepTime[12] := 1, [1].StepTime[13] := 3, [1].StepTime[14] := 3, [1].StepTime[15] := 10, [1].StepTime[16] := 20, [1].StepTime[17] := 1, [1].StepTime[18] := 1, [1].StepTime[19] := 3, [1].StepTime[20] := 15, [1].StepTime[21] := 50, [1].StepTime[22] := 1, [1].StepTime[23] := 1, [1].StepTime[24] := 3, [1].StepTime[25] := 10, [1].StepTime[26] := 20, [1].StepTime[27] := 1, [1].StepTime[28] := 1, [1].StepTime[29] := 20, [1].StepTime[30] := 40, [1].StepTime[31] := 1, [1].StepTime[32] := 1, [1].StepTime[33] := 10, [1].StepTime[34] := 10, [1].StepTime[35] := 1,
        [1].StepTime[36] := 10, [1].StepTime[37] := 20, [1].StepTime[38] := 20, [1].StepTime[39] := 10, [1].StepTime[40] := 1, [1].Setpoint[1] := 45.0, [1].Setpoint[2] := 45.0, [1].Setpoint[3] := 45.0, [1].Setpoint[4] := 45.0, [1].Setpoint[5] := 45.0, [1].Setpoint[6] := 25.0, [1].Setpoint[7] := 42.0, [1].Setpoint[8] := 42.0, [1].Setpoint[9] := 42.0, [1].Setpoint[10] := 42.0, [1].Setpoint[11] := 42.0, [1].Setpoint[12] := 22.0, [1].Setpoint[13] := 60.0, [1].Setpoint[14] := 900.0, [1].Setpoint[15] := 300.0, [1].Setpoint[16] := 300.0, [1].Setpoint[17] := 5.0, [1].Setpoint[18] := 4.5, [1].Setpoint[19] := 30.0, [1].Setpoint[20] := 60.0, [1].Setpoint[21] := 5.0, [1].Setpoint[22] := 15.0, [1].Setpoint[23] := 300.0, [1].Setpoint[24] := 0.2, [1].Setpoint[25] := 2.0, [1].Setpoint[26] := 1.5, [1].Setpoint[27] := 60.0, [1].Setpoint[28] := 50.0, [1].Setpoint[29] := 30.0, [1].Setpoint[30] := 30.0, [1].Setpoint[31] := 300.0, [1].Setpoint[32] := 0.1, [1].Setpoint[33] := 5.0, [1].Setpoint[34] := 900.0, [1].Setpoint[37] := 70.0, [1].Setpoint[38] := 100.0, [1].Setpoint[39] := 110.0, [1].Setpoint[40] := 30.0, [1].Setpoint[41] := 60.0, [1].Setpoint[42] := 900.0, [1].Setpoint[43] := 3000.0, [1].Setpoint[44] := 300.0, [1].Setpoint[45] := 195.0, [1].Setpoint[46] := 10.0, [1].Setpoint[47] := 150.0, [1].Setpoint[48] := 190.0, [1].Setpoint[49] := 60.0, [1].Setpoint[50] := 60.0, [1].Setpoint[51] := 80.0, [1].Setpoint[52] := 190.0, [1].Setpoint[53] := 50.0, [1].Setpoint[54] := 85.0, [1].Setpoint[55] := 40.0, [1].Setpoint[56] := 25.0, [1].Setpoint[57] := 10.0,
        [1].Setpoint[58] := 4.0, [1].Setpoint[61] := 5.0, [1].Setpoint[62] := 1.0, [1].Setpoint[65] := 100.0, [1].Setpoint[66] := 15.0, [1].Setpoint[67] := 50.0, [1].Setpoint[68] := 5.0, [1].Setpoint[69] := 60.0, [1].Setpoint[70] := 20.0, [1].Setpoint[71] := 60.0, [1].Setpoint[72] := 2.0, [1].Setpoint[73] := 120.0, [1].Setpoint[74] := 20.0, [1].Setpoint[75] := 120.0, [1].Setpoint[76] := 20.0, [1].Setpoint[77] := 40.0, [1].Setpoint[78] := 15.0, [1].Setpoint[79] := 30.0, [1].Setpoint[80] := 5.0, [1].Setpoint[81] := 45.0, [1].Setpoint[82] := 30.0, [1].Setpoint[83] := 5.0, [1].Setpoint[85] := 5.5, [1].Setpoint[86] := 10.5, [1].Setpoint[92] := 75.0, [1].Setpoint[93] := 90.0, [1].Setpoint[94] := 5.0, [1].Setpoint[95] := 110.0, [1].Setpoint[96] := 10.0, [1].Name := 'TANK WASH W/DIP TUBES CYCLE', [2].OpCode[1] := 50, [2].OpCode[2] := 5, [2].OpCode[3] := 52, [2].OpCode[4] := 12, [2].OpCode[5] := 11, [2].OpCode[6] := 65, [2].OpCode[7] := 41, [2].OpCode[8] := 5, [2].OpCode[9] := 33, [2].OpCode[10] := 16, [2].OpCode[11] := 15, [2].OpCode[12] := 67, [2].OpCode[13] := 38, [2].OpCode[14] := 41, [2].OpCode[15] := 2, [2].OpCode[16] := 8, [2].OpCode[17] := 51, [2].OpCode[18] := 5, [2].OpCode[19] := 6, [2].OpCode[20] := 28, [2].OpCode[21] := 27, [2].OpCode[22] := 66, [2].OpCode[23] := 38, [2].OpCode[24] := 41, [2].OpCode[25] := 2, [2].OpCode[26] := 8, [2].OpCode[27] := 49, [2].OpCode[28] := 5, [2].OpCode[29] := 24, [2].OpCode[30] := 23,
        [2].OpCode[31] := 66, [2].OpCode[32] := 5, [2].OpCode[33] := 32, [2].OpCode[34] := 31, [2].OpCode[35] := 69, [2].OpCode[36] := 2, [2].OpCode[37] := 44, [2].OpCode[38] := 45, [2].OpCode[39] := 4, [2].OpCode[40] := 1, [2].StepTime[1] := 1, [2].StepTime[2] := 1, [2].StepTime[3] := 1, [2].StepTime[4] := 10, [2].StepTime[5] := 70, [2].StepTime[6] := 1, [2].StepTime[7] := 3, [2].StepTime[8] := 1, [2].StepTime[9] := 30, [2].StepTime[10] := 50, [2].StepTime[11] := 150, [2].StepTime[12] := 1, [2].StepTime[13] := 3, [2].StepTime[14] := 3, [2].StepTime[15] := 10, [2].StepTime[16] := 20, [2].StepTime[17] := 1, [2].StepTime[18] := 1, [2].StepTime[19] := 3, [2].StepTime[20] := 15, [2].StepTime[21] := 50, [2].StepTime[22] := 1, [2].StepTime[23] := 1, [2].StepTime[24] := 3, [2].StepTime[25] := 10, [2].StepTime[26] := 20, [2].StepTime[27] := 1, [2].StepTime[28] := 1, [2].StepTime[29] := 20, [2].StepTime[30] := 40, [2].StepTime[31] := 1, [2].StepTime[32] := 1, [2].StepTime[33] := 10, [2].StepTime[34] := 10, [2].StepTime[35] := 1, [2].StepTime[36] := 10, [2].StepTime[37] := 20, [2].StepTime[38] := 20, [2].StepTime[39] := 10, [2].StepTime[40] := 1, [2].Setpoint[1] := 45.0, [2].Setpoint[2] := 45.0, [2].Setpoint[3] := 45.0, [2].Setpoint[4] := 45.0, [2].Setpoint[5] := 45.0, [2].Setpoint[6] := 25.0, [2].Setpoint[7] := 42.0, [2].Setpoint[8] := 42.0, [2].Setpoint[9] := 42.0, [2].Setpoint[10] := 42.0,
        [2].Setpoint[11] := 42.0, [2].Setpoint[12] := 22.0, [2].Setpoint[13] := 60.0, [2].Setpoint[14] := 900.0, [2].Setpoint[15] := 300.0, [2].Setpoint[16] := 300.0, [2].Setpoint[17] := 5.0, [2].Setpoint[18] := 4.5, [2].Setpoint[19] := 30.0, [2].Setpoint[20] := 60.0, [2].Setpoint[21] := 5.0, [2].Setpoint[22] := 15.0, [2].Setpoint[23] := 300.0, [2].Setpoint[24] := 0.2, [2].Setpoint[25] := 2.0, [2].Setpoint[26] := 1.5, [2].Setpoint[27] := 60.0, [2].Setpoint[28] := 50.0, [2].Setpoint[29] := 30.0, [2].Setpoint[30] := 30.0, [2].Setpoint[31] := 300.0, [2].Setpoint[32] := 0.1, [2].Setpoint[33] := 5.0, [2].Setpoint[34] := 900.0, [2].Setpoint[37] := 70.0, [2].Setpoint[38] := 100.0, [2].Setpoint[39] := 110.0, [2].Setpoint[40] := 30.0, [2].Setpoint[41] := 60.0, [2].Setpoint[42] := 900.0, [2].Setpoint[43] := 3000.0, [2].Setpoint[44] := 300.0, [2].Setpoint[45] := 195.0, [2].Setpoint[46] := 10.0, [2].Setpoint[47] := 150.0, [2].Setpoint[48] := 190.0, [2].Setpoint[49] := 60.0, [2].Setpoint[50] := 60.0, [2].Setpoint[51] := 80.0, [2].Setpoint[52] := 190.0, [2].Setpoint[53] := 50.0, [2].Setpoint[54] := 85.0, [2].Setpoint[55] := 40.0, [2].Setpoint[56] := 25.0, [2].Setpoint[57] := 10.0, [2].Setpoint[58] := 4.0, [2].Setpoint[61] := 5.0, [2].Setpoint[62] := 1.0, [2].Setpoint[65] := 100.0, [2].Setpoint[66] := 15.0, [2].Setpoint[67] := 50.0, [2].Setpoint[68] := 5.0, [2].Setpoint[69] := 60.0, [2].Setpoint[70] := 20.0, [2].Setpoint[71] := 60.0, [2].Setpoint[72] := 2.0, [2].Setpoint[73] := 120.0, [2].Setpoint[74] := 20.0, [2].Setpoint[75] := 120.0, [2].Setpoint[76] := 20.0,
        [2].Setpoint[77] := 40.0, [2].Setpoint[78] := 15.0, [2].Setpoint[79] := 30.0, [2].Setpoint[80] := 5.0, [2].Setpoint[81] := 45.0, [2].Setpoint[82] := 30.0, [2].Setpoint[83] := 5.0, [2].Setpoint[85] := 5.5, [2].Setpoint[86] := 10.5, [2].Setpoint[92] := 75.0, [2].Setpoint[93] := 90.0, [2].Setpoint[94] := 5.0, [2].Setpoint[95] := 110.0, [2].Setpoint[96] := 10.0, [2].Name := 'TANK WASH W/DIP TUBES CYCLE #2', [3].OpCode[1] := 50, [3].OpCode[2] := 5, [3].OpCode[3] := 52, [3].OpCode[4] := 9, [3].OpCode[5] := 10, [3].OpCode[6] := 65, [3].OpCode[7] := 40, [3].OpCode[8] := 5, [3].OpCode[9] := 33, [3].OpCode[10] := 13, [3].OpCode[11] := 14, [3].OpCode[12] := 67, [3].OpCode[13] := 37, [3].OpCode[14] := 40, [3].OpCode[15] := 2, [3].OpCode[16] := 8, [3].OpCode[17] := 51, [3].OpCode[18] := 5, [3].OpCode[19] := 6, [3].OpCode[20] := 25, [3].OpCode[21] := 26, [3].OpCode[22] := 66, [3].OpCode[23] := 40, [3].OpCode[24] := 2, [3].OpCode[25] := 8, [3].OpCode[26] := 49, [3].OpCode[27] := 5, [3].OpCode[28] := 21, [3].OpCode[29] := 22, [3].OpCode[30] := 40, [3].OpCode[31] := 5, [3].OpCode[32] := 29, [3].OpCode[33] := 30, [3].OpCode[34] := 69, [3].OpCode[35] := 40, [3].OpCode[36] := 46, [3].OpCode[37] := 47, [3].OpCode[38] := 43, [3].OpCode[39] := 2, [3].OpCode[40] := 35, [3].OpCode[41] := 36, [3].OpCode[42] := 1, [3].StepTime[1] := 1, [3].StepTime[2] := 1, [3].StepTime[3] := 1,
        [3].StepTime[4] := 15, [3].StepTime[5] := 6, [3].StepTime[6] := 1, [3].StepTime[7] := 3, [3].StepTime[8] := 1, [3].StepTime[9] := 30, [3].StepTime[10] := 100, [3].StepTime[11] := 100, [3].StepTime[12] := 1, [3].StepTime[13] := 1, [3].StepTime[14] := 3, [3].StepTime[15] := 10, [3].StepTime[16] := 20, [3].StepTime[17] := 1, [3].StepTime[18] := 1, [3].StepTime[19] := 3, [3].StepTime[20] := 15, [3].StepTime[21] := 15, [3].StepTime[22] := 1, [3].StepTime[23] := 3, [3].StepTime[24] := 10, [3].StepTime[25] := 20, [3].StepTime[26] := 10, [3].StepTime[27] := 1, [3].StepTime[28] := 10, [3].StepTime[29] := 10, [3].StepTime[30] := 3, [3].StepTime[31] := 1, [3].StepTime[32] := 5, [3].StepTime[33] := 5, [3].StepTime[34] := 1, [3].StepTime[35] := 3, [3].StepTime[36] := 5, [3].StepTime[37] := 5, [3].StepTime[38] := 3, [3].StepTime[39] := 10, [3].StepTime[40] := 200, [3].StepTime[41] := 30, [3].StepTime[42] := 1, [3].Setpoint[1] := 45.0, [3].Setpoint[2] := 45.0, [3].Setpoint[3] := 45.0, [3].Setpoint[4] := 45.0, [3].Setpoint[5] := 45.0, [3].Setpoint[6] := 25.0, [3].Setpoint[7] := 42.0, [3].Setpoint[8] := 42.0, [3].Setpoint[9] := 42.0, [3].Setpoint[10] := 42.0, [3].Setpoint[11] := 42.0, [3].Setpoint[12] := 22.0, [3].Setpoint[13] := 60.0, [3].Setpoint[14] := 900.0, [3].Setpoint[15] := 300.0, [3].Setpoint[16] := 300.0, [3].Setpoint[17] := 5.0, [3].Setpoint[18] := 4.5, [3].Setpoint[19] := 45.0, [3].Setpoint[20] := 60.0, [3].Setpoint[21] := 5.0,
        [3].Setpoint[22] := 15.0, [3].Setpoint[23] := 300.0, [3].Setpoint[24] := 0.2, [3].Setpoint[25] := 10.0, [3].Setpoint[26] := 9.0, [3].Setpoint[27] := 30.0, [3].Setpoint[28] := 50.0, [3].Setpoint[29] := 3.0, [3].Setpoint[30] := 17.0, [3].Setpoint[31] := 300.0, [3].Setpoint[32] := 2.0, [3].Setpoint[33] := 5.0, [3].Setpoint[34] := 900.0, [3].Setpoint[37] := 50.0, [3].Setpoint[38] := 75.0, [3].Setpoint[39] := 100.0, [3].Setpoint[40] := 30.0, [3].Setpoint[41] := 60.0, [3].Setpoint[42] := 900.0, [3].Setpoint[43] := 3000.0, [3].Setpoint[44] := 300.0, [3].Setpoint[45] := 195.0, [3].Setpoint[46] := 10.0, [3].Setpoint[47] := 186.0, [3].Setpoint[48] := 190.0, [3].Setpoint[49] := 80.0, [3].Setpoint[50] := 80.0, [3].Setpoint[51] := 80.0, [3].Setpoint[52] := 185.0, [3].Setpoint[53] := 50.0, [3].Setpoint[54] := 85.0, [3].Setpoint[55] := 100.0, [3].Setpoint[56] := 60.0, [3].Setpoint[57] := 90.0, [3].Setpoint[58] := 4.0, [3].Setpoint[62] := 1.0, [3].Setpoint[65] := 80.0, [3].Setpoint[66] := 15.0, [3].Setpoint[67] := 65.0, [3].Setpoint[68] := 5.0, [3].Setpoint[69] := 100.0, [3].Setpoint[70] := 15.0, [3].Setpoint[71] := 100.0, [3].Setpoint[72] := 15.0, [3].Setpoint[73] := 120.0, [3].Setpoint[74] := 20.0, [3].Setpoint[75] := 120.0, [3].Setpoint[76] := 20.0, [3].Setpoint[77] := 100.0, [3].Setpoint[78] := 15.0, [3].Setpoint[79] := 100.0, [3].Setpoint[80] := 15.0, [3].Setpoint[81] := 47.0, [3].Setpoint[82] := 20.0, [3].Setpoint[83] := 5.0, [3].Setpoint[84] := 1.0, [3].Setpoint[85] := 5.5, [3].Setpoint[86] := 10.5, [3].Setpoint[92] := 75.0, [3].Setpoint[93] := 90.0,
        [3].Setpoint[94] := 5.0, [3].Setpoint[95] := 110.0, [3].Setpoint[96] := 10.0, [3].Name := 'WASH CHAMBER WASH CYCLE POLY/GLASSWARE', [4].OpCode[1] := 50, [4].OpCode[2] := 5, [4].OpCode[3] := 52, [4].OpCode[4] := 9, [4].OpCode[5] := 10, [4].OpCode[6] := 65, [4].OpCode[7] := 40, [4].OpCode[8] := 5, [4].OpCode[9] := 33, [4].OpCode[10] := 13, [4].OpCode[11] := 14, [4].OpCode[12] := 67, [4].OpCode[13] := 37, [4].OpCode[14] := 40, [4].OpCode[15] := 2, [4].OpCode[16] := 8, [4].OpCode[17] := 51, [4].OpCode[18] := 5, [4].OpCode[19] := 6, [4].OpCode[20] := 25, [4].OpCode[21] := 26, [4].OpCode[22] := 66, [4].OpCode[23] := 40, [4].OpCode[24] := 2, [4].OpCode[25] := 8, [4].OpCode[26] := 49, [4].OpCode[27] := 5, [4].OpCode[28] := 21, [4].OpCode[29] := 22, [4].OpCode[30] := 40, [4].OpCode[31] := 5, [4].OpCode[32] := 29, [4].OpCode[33] := 30, [4].OpCode[34] := 69, [4].OpCode[35] := 40, [4].OpCode[36] := 46, [4].OpCode[37] := 47, [4].OpCode[38] := 43, [4].OpCode[39] := 2, [4].OpCode[40] := 35, [4].OpCode[41] := 36, [4].OpCode[42] := 1, [4].StepTime[1] := 1, [4].StepTime[2] := 1, [4].StepTime[3] := 1, [4].StepTime[4] := 15, [4].StepTime[5] := 6, [4].StepTime[6] := 1, [4].StepTime[7] := 3, [4].StepTime[8] := 1, [4].StepTime[9] := 30, [4].StepTime[10] := 100, [4].StepTime[11] := 100, [4].StepTime[12] := 1, [4].StepTime[13] := 1, [4].StepTime[14] := 3,
        [4].StepTime[15] := 10, [4].StepTime[16] := 20, [4].StepTime[17] := 1, [4].StepTime[18] := 1, [4].StepTime[19] := 3, [4].StepTime[20] := 15, [4].StepTime[21] := 15, [4].StepTime[22] := 1, [4].StepTime[23] := 3, [4].StepTime[24] := 10, [4].StepTime[25] := 20, [4].StepTime[26] := 10, [4].StepTime[27] := 1, [4].StepTime[28] := 10, [4].StepTime[29] := 10, [4].StepTime[30] := 3, [4].StepTime[31] := 1, [4].StepTime[32] := 5, [4].StepTime[33] := 5, [4].StepTime[34] := 1, [4].StepTime[35] := 3, [4].StepTime[36] := 5, [4].StepTime[37] := 5, [4].StepTime[38] := 3, [4].StepTime[39] := 10, [4].StepTime[40] := 200, [4].StepTime[41] := 30, [4].StepTime[42] := 1, [4].Setpoint[1] := 45.0, [4].Setpoint[2] := 45.0, [4].Setpoint[3] := 45.0, [4].Setpoint[4] := 45.0, [4].Setpoint[5] := 45.0, [4].Setpoint[6] := 25.0, [4].Setpoint[7] := 42.0, [4].Setpoint[8] := 42.0, [4].Setpoint[9] := 42.0, [4].Setpoint[10] := 42.0, [4].Setpoint[11] := 42.0, [4].Setpoint[12] := 22.0, [4].Setpoint[13] := 60.0, [4].Setpoint[14] := 900.0, [4].Setpoint[15] := 300.0, [4].Setpoint[16] := 300.0, [4].Setpoint[17] := 5.0, [4].Setpoint[18] := 4.5, [4].Setpoint[19] := 45.0, [4].Setpoint[20] := 60.0, [4].Setpoint[21] := 5.0, [4].Setpoint[22] := 15.0, [4].Setpoint[23] := 300.0, [4].Setpoint[24] := 0.2, [4].Setpoint[25] := 10.0, [4].Setpoint[26] := 9.0, [4].Setpoint[27] := 30.0, [4].Setpoint[28] := 50.0, [4].Setpoint[29] := 3.0, [4].Setpoint[30] := 17.0, [4].Setpoint[31] := 300.0, [4].Setpoint[32] := 2.0,
        [4].Setpoint[33] := 5.0, [4].Setpoint[34] := 900.0, [4].Setpoint[37] := 50.0, [4].Setpoint[38] := 75.0, [4].Setpoint[39] := 100.0, [4].Setpoint[40] := 30.0, [4].Setpoint[41] := 60.0, [4].Setpoint[42] := 900.0, [4].Setpoint[43] := 3000.0, [4].Setpoint[44] := 300.0, [4].Setpoint[45] := 195.0, [4].Setpoint[46] := 10.0, [4].Setpoint[47] := 186.0, [4].Setpoint[48] := 190.0, [4].Setpoint[49] := 80.0, [4].Setpoint[50] := 80.0, [4].Setpoint[51] := 80.0, [4].Setpoint[52] := 185.0, [4].Setpoint[53] := 50.0, [4].Setpoint[54] := 85.0, [4].Setpoint[55] := 100.0, [4].Setpoint[56] := 60.0, [4].Setpoint[57] := 90.0, [4].Setpoint[58] := 4.0, [4].Setpoint[62] := 1.0, [4].Setpoint[65] := 80.0, [4].Setpoint[66] := 15.0, [4].Setpoint[67] := 65.0, [4].Setpoint[68] := 5.0, [4].Setpoint[69] := 100.0, [4].Setpoint[70] := 15.0, [4].Setpoint[71] := 100.0, [4].Setpoint[72] := 15.0, [4].Setpoint[73] := 120.0, [4].Setpoint[74] := 20.0, [4].Setpoint[75] := 120.0, [4].Setpoint[76] := 20.0, [4].Setpoint[77] := 100.0, [4].Setpoint[78] := 15.0, [4].Setpoint[79] := 100.0, [4].Setpoint[80] := 15.0, [4].Setpoint[81] := 47.0, [4].Setpoint[82] := 20.0, [4].Setpoint[83] := 5.0, [4].Setpoint[84] := 1.0, [4].Setpoint[85] := 5.5, [4].Setpoint[86] := 10.5, [4].Setpoint[92] := 75.0, [4].Setpoint[93] := 90.0, [4].Setpoint[94] := 5.0, [4].Setpoint[95] := 110.0, [4].Setpoint[96] := 10.0, [4].Name := 'WASH CHAMBER WAS CYCLE PROCESS PARTS', [5].OpCode[1] := 50, [5].OpCode[2] := 5, [5].OpCode[3] := 52, [5].OpCode[4] := 12, [5].OpCode[5] := 65, [5].OpCode[6] := 5, [5].OpCode[7] := 33,
        [5].OpCode[8] := 16, [5].OpCode[9] := 67, [5].OpCode[10] := 2, [5].OpCode[11] := 8, [5].OpCode[12] := 51, [5].OpCode[13] := 5, [5].OpCode[14] := 6, [5].OpCode[15] := 24, [5].OpCode[16] := 66, [5].OpCode[17] := 49, [5].OpCode[18] := 5, [5].OpCode[19] := 32, [5].OpCode[20] := 69, [5].OpCode[21] := 45, [5].OpCode[22] := 2, [5].OpCode[23] := 1, [5].StepTime[1] := 1, [5].StepTime[2] := 1, [5].StepTime[3] := 1, [5].StepTime[4] := 40, [5].StepTime[5] := 1, [5].StepTime[6] := 1, [5].StepTime[7] := 20, [5].StepTime[8] := 100, [5].StepTime[9] := 1, [5].StepTime[10] := 10, [5].StepTime[11] := 20, [5].StepTime[12] := 1, [5].StepTime[13] := 1, [5].StepTime[14] := 3, [5].StepTime[15] := 20, [5].StepTime[16] := 1, [5].StepTime[17] := 1, [5].StepTime[18] := 1, [5].StepTime[19] := 10, [5].StepTime[20] := 1, [5].StepTime[21] := 10, [5].StepTime[22] := 10, [5].StepTime[23] := 1, [5].Setpoint[1] := 45.0, [5].Setpoint[2] := 45.0, [5].Setpoint[3] := 45.0, [5].Setpoint[4] := 45.0, [5].Setpoint[5] := 45.0, [5].Setpoint[6] := 25.0, [5].Setpoint[7] := 42.0, [5].Setpoint[8] := 42.0, [5].Setpoint[9] := 42.0, [5].Setpoint[10] := 42.0, [5].Setpoint[11] := 42.0, [5].Setpoint[12] := 22.0, [5].Setpoint[13] := 60.0, [5].Setpoint[14] := 900.0, [5].Setpoint[15] := 300.0, [5].Setpoint[16] := 300.0, [5].Setpoint[17] := 5.0, [5].Setpoint[18] := 4.5, [5].Setpoint[19] := 30.0, [5].Setpoint[20] := 60.0, [5].Setpoint[21] := 5.0,
        [5].Setpoint[22] := 15.0, [5].Setpoint[23] := 300.0, [5].Setpoint[24] := 0.2, [5].Setpoint[25] := 10.0, [5].Setpoint[26] := 9.0, [5].Setpoint[27] := 10.0, [5].Setpoint[28] := 50.0, [5].Setpoint[29] := 3.0, [5].Setpoint[30] := 17.0, [5].Setpoint[31] := 300.0, [5].Setpoint[32] := 2.0, [5].Setpoint[33] := 5.0, [5].Setpoint[34] := 900.0, [5].Setpoint[37] := 70.0, [5].Setpoint[38] := 100.0, [5].Setpoint[39] := 110.0, [5].Setpoint[40] := 30.0, [5].Setpoint[41] := 60.0, [5].Setpoint[42] := 900.0, [5].Setpoint[43] := 3000.0, [5].Setpoint[44] := 300.0, [5].Setpoint[45] := 195.0, [5].Setpoint[46] := 10.0, [5].Setpoint[47] := 25.0, [5].Setpoint[48] := 190.0, [5].Setpoint[49] := 100.0, [5].Setpoint[50] := 60.0, [5].Setpoint[51] := 80.0, [5].Setpoint[52] := 185.0, [5].Setpoint[53] := 50.0, [5].Setpoint[54] := 85.0, [5].Setpoint[55] := 40.0, [5].Setpoint[56] := 60.0, [5].Setpoint[57] := 43.0, [5].Setpoint[58] := 4.0, [5].Setpoint[61] := 10.0, [5].Setpoint[62] := 1.0, [5].Setpoint[65] := 100.0, [5].Setpoint[66] := 15.0, [5].Setpoint[67] := 50.0, [5].Setpoint[68] := 5.0, [5].Setpoint[69] := 100.0, [5].Setpoint[70] := 15.0, [5].Setpoint[71] := 40.0, [5].Setpoint[72] := 2.0, [5].Setpoint[73] := 120.0, [5].Setpoint[74] := 20.0, [5].Setpoint[75] := 120.0, [5].Setpoint[76] := 20.0, [5].Setpoint[77] := 100.0, [5].Setpoint[78] := 15.0, [5].Setpoint[79] := 60.0, [5].Setpoint[80] := 30.0, [5].Setpoint[81] := 45.0, [5].Setpoint[82] := 30.0, [5].Setpoint[83] := 5.0, [5].Setpoint[85] := 5.5, [5].Setpoint[86] := 10.5, [5].Setpoint[92] := 75.0, [5].Setpoint[93] := 90.0,
        [5].Setpoint[94] := 5.0, [5].Setpoint[95] := 110.0, [5].Setpoint[96] := 10.0, [5].Name := 'PROCESS HOSES', [6].Setpoint[1] := 55.0, [6].Setpoint[2] := 65.0, [6].Setpoint[3] := 60.0, [6].Setpoint[4] := 45.0, [6].Setpoint[5] := 65.0, [6].Setpoint[6] := 25.0, [6].Setpoint[7] := 53.0, [6].Setpoint[8] := 63.0, [6].Setpoint[9] := 57.0, [6].Setpoint[10] := 43.0, [6].Setpoint[11] := 63.0, [6].Setpoint[12] := 22.0, [6].Setpoint[13] := 85.0, [6].Setpoint[14] := 900.0, [6].Setpoint[15] := 300.0, [6].Setpoint[16] := 300.0, [6].Setpoint[17] := 15.0, [6].Setpoint[18] := 14.0, [6].Setpoint[19] := 15.0, [6].Setpoint[20] := 45.0, [6].Setpoint[21] := 5.0, [6].Setpoint[22] := 15.0, [6].Setpoint[23] := 300.0, [6].Setpoint[24] := 2.0, [6].Setpoint[25] := 10.0, [6].Setpoint[26] := 9.0, [6].Setpoint[27] := 10.0, [6].Setpoint[28] := 50.0, [6].Setpoint[29] := 3.0, [6].Setpoint[30] := 17.0, [6].Setpoint[31] := 300.0, [6].Setpoint[32] := 2.0, [6].Setpoint[33] := 2.0, [6].Setpoint[34] := 900.0, [6].Setpoint[37] := 70.0, [6].Setpoint[38] := 90.0, [6].Setpoint[39] := 110.0, [6].Setpoint[40] := 30.0, [6].Setpoint[41] := 60.0, [6].Setpoint[42] := 60.0, [6].Setpoint[43] := 3000.0, [6].Setpoint[44] := 300.0, [6].Setpoint[45] := 190.0, [6].Setpoint[46] := 10.0, [6].Setpoint[47] := 25.0, [6].Setpoint[48] := 150.0, [6].Setpoint[49] := 125.0, [6].Setpoint[50] := 100.0, [6].Setpoint[51] := 80.0, [6].Setpoint[52] := 100.0, [6].Setpoint[53] := 50.0, [6].Setpoint[54] := 85.0, [6].Setpoint[55] := 40.0, [6].Setpoint[56] := 60.0, [6].Setpoint[57] := 90.0, [6].Setpoint[58] := 4.0,
        [6].Setpoint[61] := 10.0, [6].Setpoint[62] := 1.0, [6].Setpoint[65] := 100.0, [6].Setpoint[66] := 15.0, [6].Setpoint[67] := 50.0, [6].Setpoint[68] := 5.0, [6].Setpoint[69] := 100.0, [6].Setpoint[70] := 15.0, [6].Setpoint[71] := 100.0, [6].Setpoint[72] := 15.0, [6].Setpoint[73] := 120.0, [6].Setpoint[74] := 20.0, [6].Setpoint[75] := 120.0, [6].Setpoint[76] := 20.0, [6].Setpoint[77] := 100.0, [6].Setpoint[78] := 15.0, [6].Setpoint[79] := 100.0, [6].Setpoint[80] := 15.0, [6].Setpoint[81] := 45.0, [6].Setpoint[82] := 30.0, [6].Setpoint[83] := 5.0, [6].Setpoint[84] := 1.0, [6].Setpoint[85] := 5.0, [6].Setpoint[86] := 9.0, [6].Setpoint[92] := 75.0, [6].Setpoint[93] := 90.0, [6].Setpoint[94] := 5.0, [6].Setpoint[95] := 110.0, [6].Setpoint[96] := 10.0, [6].Name := 'RECIPE #6', [7].Setpoint[1] := 55.0, [7].Setpoint[2] := 65.0, [7].Setpoint[3] := 60.0, [7].Setpoint[4] := 45.0, [7].Setpoint[5] := 65.0, [7].Setpoint[6] := 25.0, [7].Setpoint[7] := 53.0, [7].Setpoint[8] := 63.0, [7].Setpoint[9] := 57.0, [7].Setpoint[10] := 43.0, [7].Setpoint[11] := 63.0, [7].Setpoint[12] := 22.0, [7].Setpoint[13] := 85.0, [7].Setpoint[14] := 900.0, [7].Setpoint[15] := 300.0, [7].Setpoint[16] := 300.0, [7].Setpoint[17] := 15.0, [7].Setpoint[18] := 14.0, [7].Setpoint[19] := 15.0, [7].Setpoint[20] := 45.0, [7].Setpoint[21] := 5.0, [7].Setpoint[22] := 15.0, [7].Setpoint[23] := 300.0, [7].Setpoint[24] := 2.0, [7].Setpoint[25] := 10.0, [7].Setpoint[26] := 9.0, [7].Setpoint[27] := 10.0, [7].Setpoint[28] := 50.0, [7].Setpoint[29] := 3.0, [7].Setpoint[30] := 17.0,
        [7].Setpoint[31] := 300.0, [7].Setpoint[32] := 2.0, [7].Setpoint[33] := 2.0, [7].Setpoint[34] := 900.0, [7].Setpoint[37] := 70.0, [7].Setpoint[38] := 100.0, [7].Setpoint[39] := 110.0, [7].Setpoint[40] := 30.0, [7].Setpoint[41] := 60.0, [7].Setpoint[42] := 60.0, [7].Setpoint[43] := 3000.0, [7].Setpoint[44] := 300.0, [7].Setpoint[45] := 185.0, [7].Setpoint[46] := 10.0, [7].Setpoint[47] := 25.0, [7].Setpoint[48] := 150.0, [7].Setpoint[49] := 125.0, [7].Setpoint[50] := 100.0, [7].Setpoint[51] := 80.0, [7].Setpoint[52] := 100.0, [7].Setpoint[53] := 50.0, [7].Setpoint[54] := 85.0, [7].Setpoint[55] := 40.0, [7].Setpoint[56] := 60.0, [7].Setpoint[57] := 90.0, [7].Setpoint[58] := 4.0, [7].Setpoint[61] := 10.0, [7].Setpoint[62] := 1.0, [7].Setpoint[65] := 100.0, [7].Setpoint[66] := 15.0, [7].Setpoint[67] := 50.0, [7].Setpoint[68] := 5.0, [7].Setpoint[69] := 100.0, [7].Setpoint[70] := 15.0, [7].Setpoint[71] := 100.0, [7].Setpoint[72] := 15.0, [7].Setpoint[73] := 120.0, [7].Setpoint[74] := 20.0, [7].Setpoint[75] := 120.0, [7].Setpoint[76] := 20.0, [7].Setpoint[77] := 100.0, [7].Setpoint[78] := 15.0, [7].Setpoint[79] := 100.0, [7].Setpoint[80] := 15.0, [7].Setpoint[81] := 45.0, [7].Setpoint[82] := 30.0, [7].Setpoint[83] := 5.0, [7].Setpoint[85] := 5.0, [7].Setpoint[86] := 9.0, [7].Setpoint[92] := 75.0, [7].Setpoint[93] := 90.0, [7].Setpoint[94] := 5.0, [7].Setpoint[95] := 110.0, [7].Setpoint[96] := 10.0, [7].Name := 'RECIPE #7', [8].Setpoint[1] := 55.0, [8].Setpoint[2] := 65.0, [8].Setpoint[3] := 60.0, [8].Setpoint[4] := 45.0, [8].Setpoint[5] := 65.0,
        [8].Setpoint[6] := 25.0, [8].Setpoint[7] := 53.0, [8].Setpoint[8] := 63.0, [8].Setpoint[9] := 57.0, [8].Setpoint[10] := 43.0, [8].Setpoint[11] := 63.0, [8].Setpoint[12] := 22.0, [8].Setpoint[13] := 85.0, [8].Setpoint[14] := 900.0, [8].Setpoint[15] := 300.0, [8].Setpoint[16] := 300.0, [8].Setpoint[17] := 15.0, [8].Setpoint[18] := 14.0, [8].Setpoint[19] := 15.0, [8].Setpoint[20] := 45.0, [8].Setpoint[21] := 5.0, [8].Setpoint[22] := 15.0, [8].Setpoint[23] := 300.0, [8].Setpoint[24] := 2.0, [8].Setpoint[25] := 10.0, [8].Setpoint[26] := 9.0, [8].Setpoint[27] := 10.0, [8].Setpoint[28] := 50.0, [8].Setpoint[29] := 3.0, [8].Setpoint[30] := 17.0, [8].Setpoint[31] := 300.0, [8].Setpoint[32] := 2.0, [8].Setpoint[33] := 2.0, [8].Setpoint[34] := 900.0, [8].Setpoint[37] := 70.0, [8].Setpoint[38] := 100.0, [8].Setpoint[39] := 110.0, [8].Setpoint[40] := 30.0, [8].Setpoint[41] := 60.0, [8].Setpoint[42] := 60.0, [8].Setpoint[43] := 3000.0, [8].Setpoint[44] := 300.0, [8].Setpoint[45] := 185.0, [8].Setpoint[46] := 10.0, [8].Setpoint[47] := 25.0, [8].Setpoint[48] := 150.0, [8].Setpoint[49] := 125.0, [8].Setpoint[50] := 100.0, [8].Setpoint[51] := 80.0, [8].Setpoint[52] := 100.0, [8].Setpoint[53] := 50.0, [8].Setpoint[54] := 85.0, [8].Setpoint[55] := 40.0, [8].Setpoint[56] := 60.0, [8].Setpoint[57] := 90.0, [8].Setpoint[58] := 4.0, [8].Setpoint[61] := 10.0, [8].Setpoint[62] := 1.0, [8].Setpoint[65] := 100.0, [8].Setpoint[66] := 15.0, [8].Setpoint[67] := 50.0, [8].Setpoint[68] := 5.0, [8].Setpoint[69] := 100.0, [8].Setpoint[70] := 15.0, [8].Setpoint[71] := 100.0,
        [8].Setpoint[72] := 15.0, [8].Setpoint[73] := 120.0, [8].Setpoint[74] := 20.0, [8].Setpoint[75] := 120.0, [8].Setpoint[76] := 20.0, [8].Setpoint[77] := 100.0, [8].Setpoint[78] := 15.0, [8].Setpoint[79] := 100.0, [8].Setpoint[80] := 15.0, [8].Setpoint[81] := 45.0, [8].Setpoint[82] := 30.0, [8].Setpoint[83] := 5.0, [8].Setpoint[85] := 5.0, [8].Setpoint[86] := 9.0, [8].Setpoint[92] := 75.0, [8].Setpoint[93] := 90.0, [8].Setpoint[94] := 5.0, [8].Setpoint[95] := 110.0, [8].Setpoint[96] := 10.0, [8].Name := 'RECIPE #8', [9].Setpoint[1] := 55.0, [9].Setpoint[2] := 65.0, [9].Setpoint[3] := 60.0, [9].Setpoint[4] := 45.0, [9].Setpoint[5] := 65.0, [9].Setpoint[6] := 25.0, [9].Setpoint[7] := 53.0, [9].Setpoint[8] := 63.0, [9].Setpoint[9] := 57.0, [9].Setpoint[10] := 43.0, [9].Setpoint[11] := 63.0, [9].Setpoint[12] := 22.0, [9].Setpoint[13] := 85.0, [9].Setpoint[14] := 900.0, [9].Setpoint[15] := 300.0, [9].Setpoint[16] := 300.0, [9].Setpoint[17] := 15.0, [9].Setpoint[18] := 14.0, [9].Setpoint[19] := 15.0, [9].Setpoint[20] := 45.0, [9].Setpoint[21] := 5.0, [9].Setpoint[22] := 15.0, [9].Setpoint[23] := 300.0, [9].Setpoint[24] := 2.0, [9].Setpoint[25] := 10.0, [9].Setpoint[26] := 9.0, [9].Setpoint[27] := 10.0, [9].Setpoint[28] := 50.0, [9].Setpoint[29] := 3.0, [9].Setpoint[30] := 17.0, [9].Setpoint[31] := 300.0, [9].Setpoint[32] := 2.0, [9].Setpoint[33] := 2.0, [9].Setpoint[34] := 900.0, [9].Setpoint[37] := 70.0, [9].Setpoint[38] := 100.0, [9].Setpoint[39] := 110.0, [9].Setpoint[40] := 30.0, [9].Setpoint[41] := 60.0, [9].Setpoint[42] := 60.0,
        [9].Setpoint[43] := 3000.0, [9].Setpoint[44] := 300.0, [9].Setpoint[45] := 185.0, [9].Setpoint[46] := 10.0, [9].Setpoint[47] := 25.0, [9].Setpoint[48] := 150.0, [9].Setpoint[49] := 125.0, [9].Setpoint[50] := 100.0, [9].Setpoint[51] := 80.0, [9].Setpoint[52] := 100.0, [9].Setpoint[53] := 50.0, [9].Setpoint[54] := 85.0, [9].Setpoint[55] := 40.0, [9].Setpoint[56] := 60.0, [9].Setpoint[57] := 90.0, [9].Setpoint[58] := 4.0, [9].Setpoint[61] := 10.0, [9].Setpoint[62] := 1.0, [9].Setpoint[65] := 100.0, [9].Setpoint[66] := 15.0, [9].Setpoint[67] := 50.0, [9].Setpoint[68] := 5.0, [9].Setpoint[69] := 100.0, [9].Setpoint[70] := 15.0, [9].Setpoint[71] := 100.0, [9].Setpoint[72] := 15.0, [9].Setpoint[73] := 120.0, [9].Setpoint[74] := 20.0, [9].Setpoint[75] := 120.0, [9].Setpoint[76] := 20.0, [9].Setpoint[77] := 100.0, [9].Setpoint[78] := 15.0, [9].Setpoint[79] := 100.0, [9].Setpoint[80] := 15.0, [9].Setpoint[81] := 45.0, [9].Setpoint[82] := 30.0, [9].Setpoint[83] := 5.0, [9].Setpoint[85] := 5.0, [9].Setpoint[86] := 9.0, [9].Setpoint[92] := 75.0, [9].Setpoint[93] := 90.0, [9].Setpoint[94] := 5.0, [9].Setpoint[95] := 110.0, [9].Setpoint[96] := 10.0, [9].Name := 'RECIPE #9', [10].Setpoint[1] := 45.0, [10].Setpoint[2] := 45.0, [10].Setpoint[3] := 45.0, [10].Setpoint[4] := 45.0, [10].Setpoint[5] := 45.0, [10].Setpoint[6] := 25.0, [10].Setpoint[7] := 43.0, [10].Setpoint[8] := 43.0, [10].Setpoint[9] := 43.0, [10].Setpoint[10] := 43.0, [10].Setpoint[11] := 43.0, [10].Setpoint[12] := 22.0, [10].Setpoint[13] := 60.0, [10].Setpoint[14] := 900.0, [10].Setpoint[15] := 300.0,
        [10].Setpoint[16] := 300.0, [10].Setpoint[17] := 15.0, [10].Setpoint[18] := 14.0, [10].Setpoint[19] := 15.0, [10].Setpoint[20] := 45.0, [10].Setpoint[21] := 5.0, [10].Setpoint[22] := 15.0, [10].Setpoint[23] := 300.0, [10].Setpoint[24] := 2.0, [10].Setpoint[25] := 10.0, [10].Setpoint[26] := 9.0, [10].Setpoint[27] := 10.0, [10].Setpoint[28] := 50.0, [10].Setpoint[29] := 3.0, [10].Setpoint[30] := 17.0, [10].Setpoint[31] := 300.0, [10].Setpoint[32] := 2.0, [10].Setpoint[33] := 2.0, [10].Setpoint[34] := 900.0, [10].Setpoint[37] := 70.0, [10].Setpoint[38] := 100.0, [10].Setpoint[39] := 110.0, [10].Setpoint[40] := 30.0, [10].Setpoint[41] := 60.0, [10].Setpoint[42] := 60.0, [10].Setpoint[43] := 3000.0, [10].Setpoint[44] := 300.0, [10].Setpoint[45] := 200.0, [10].Setpoint[46] := 10.0, [10].Setpoint[47] := 150.0, [10].Setpoint[48] := 150.0, [10].Setpoint[49] := 150.0, [10].Setpoint[50] := 100.0, [10].Setpoint[51] := 80.0, [10].Setpoint[52] := 150.0, [10].Setpoint[53] := 50.0, [10].Setpoint[54] := 85.0, [10].Setpoint[55] := 100.0, [10].Setpoint[56] := 60.0, [10].Setpoint[57] := 90.0, [10].Setpoint[58] := 4.0, [10].Setpoint[62] := 1.0, [10].Setpoint[65] := 100.0, [10].Setpoint[66] := 15.0, [10].Setpoint[67] := 65.0, [10].Setpoint[68] := 5.0, [10].Setpoint[69] := 100.0, [10].Setpoint[70] := 15.0, [10].Setpoint[71] := 100.0, [10].Setpoint[72] := 15.0, [10].Setpoint[73] := 120.0, [10].Setpoint[74] := 20.0, [10].Setpoint[75] := 120.0, [10].Setpoint[76] := 20.0, [10].Setpoint[77] := 100.0, [10].Setpoint[78] := 15.0, [10].Setpoint[79] := 100.0, [10].Setpoint[80] := 15.0, [10].Setpoint[81] := 47.0, [10].Setpoint[82] := 30.0,
        [10].Setpoint[83] := 5.0, [10].Setpoint[84] := 1.0, [10].Setpoint[85] := 5.0, [10].Setpoint[86] := 9.0, [10].Setpoint[92] := 75.0, [10].Setpoint[93] := 90.0, [10].Setpoint[94] := 5.0, [10].Setpoint[95] := 110.0, [10].Setpoint[96] := 10.0, [10].Name := 'RECIPE #10', [11].Setpoint[1] := 55.0, [11].Setpoint[2] := 65.0, [11].Setpoint[3] := 60.0, [11].Setpoint[4] := 45.0, [11].Setpoint[5] := 65.0, [11].Setpoint[6] := 25.0, [11].Setpoint[7] := 53.0, [11].Setpoint[8] := 63.0, [11].Setpoint[9] := 57.0, [11].Setpoint[10] := 43.0, [11].Setpoint[11] := 63.0, [11].Setpoint[12] := 22.0, [11].Setpoint[13] := 85.0, [11].Setpoint[14] := 900.0, [11].Setpoint[15] := 300.0, [11].Setpoint[16] := 300.0, [11].Setpoint[17] := 15.0, [11].Setpoint[18] := 14.0, [11].Setpoint[19] := 15.0, [11].Setpoint[20] := 45.0, [11].Setpoint[21] := 5.0, [11].Setpoint[22] := 15.0, [11].Setpoint[23] := 300.0, [11].Setpoint[24] := 2.0, [11].Setpoint[25] := 10.0, [11].Setpoint[26] := 9.0, [11].Setpoint[27] := 10.0, [11].Setpoint[28] := 50.0, [11].Setpoint[29] := 3.0, [11].Setpoint[30] := 17.0, [11].Setpoint[31] := 300.0, [11].Setpoint[32] := 2.0, [11].Setpoint[33] := 2.0, [11].Setpoint[34] := 900.0, [11].Setpoint[37] := 70.0, [11].Setpoint[38] := 100.0, [11].Setpoint[39] := 110.0, [11].Setpoint[40] := 30.0, [11].Setpoint[41] := 60.0, [11].Setpoint[42] := 60.0, [11].Setpoint[43] := 3000.0, [11].Setpoint[44] := 300.0, [11].Setpoint[45] := 185.0, [11].Setpoint[46] := 10.0, [11].Setpoint[47] := 25.0, [11].Setpoint[48] := 150.0, [11].Setpoint[49] := 125.0, [11].Setpoint[50] := 100.0, [11].Setpoint[51] := 80.0, [11].Setpoint[52] := 100.0,
        [11].Setpoint[53] := 50.0, [11].Setpoint[54] := 85.0, [11].Setpoint[55] := 40.0, [11].Setpoint[56] := 60.0, [11].Setpoint[57] := 90.0, [11].Setpoint[58] := 4.0, [11].Setpoint[61] := 10.0, [11].Setpoint[62] := 1.0, [11].Setpoint[65] := 100.0, [11].Setpoint[66] := 15.0, [11].Setpoint[67] := 50.0, [11].Setpoint[68] := 5.0, [11].Setpoint[69] := 100.0, [11].Setpoint[70] := 15.0, [11].Setpoint[71] := 100.0, [11].Setpoint[72] := 15.0, [11].Setpoint[73] := 120.0, [11].Setpoint[74] := 20.0, [11].Setpoint[75] := 120.0, [11].Setpoint[76] := 20.0, [11].Setpoint[77] := 100.0, [11].Setpoint[78] := 15.0, [11].Setpoint[79] := 100.0, [11].Setpoint[80] := 15.0, [11].Setpoint[81] := 45.0, [11].Setpoint[82] := 30.0, [11].Setpoint[83] := 5.0, [11].Setpoint[85] := 5.0, [11].Setpoint[86] := 9.0, [11].Setpoint[92] := 75.0, [11].Setpoint[93] := 90.0, [11].Setpoint[94] := 5.0, [11].Setpoint[95] := 110.0, [11].Setpoint[96] := 10.0, [11].Name := 'RECIPE #11', [12].Setpoint[1] := 55.0, [12].Setpoint[2] := 65.0, [12].Setpoint[3] := 60.0, [12].Setpoint[4] := 45.0, [12].Setpoint[5] := 65.0, [12].Setpoint[6] := 25.0, [12].Setpoint[7] := 53.0, [12].Setpoint[8] := 63.0, [12].Setpoint[9] := 57.0, [12].Setpoint[10] := 43.0, [12].Setpoint[11] := 63.0, [12].Setpoint[12] := 22.0, [12].Setpoint[13] := 85.0, [12].Setpoint[14] := 900.0, [12].Setpoint[15] := 300.0, [12].Setpoint[16] := 300.0, [12].Setpoint[17] := 15.0, [12].Setpoint[18] := 14.0, [12].Setpoint[19] := 15.0, [12].Setpoint[20] := 45.0, [12].Setpoint[21] := 5.0, [12].Setpoint[22] := 15.0, [12].Setpoint[23] := 300.0, [12].Setpoint[24] := 2.0, [12].Setpoint[25] := 10.0,
        [12].Setpoint[26] := 9.0, [12].Setpoint[27] := 10.0, [12].Setpoint[28] := 50.0, [12].Setpoint[29] := 3.0, [12].Setpoint[30] := 17.0, [12].Setpoint[31] := 300.0, [12].Setpoint[32] := 2.0, [12].Setpoint[33] := 2.0, [12].Setpoint[34] := 900.0, [12].Setpoint[37] := 70.0, [12].Setpoint[38] := 100.0, [12].Setpoint[39] := 110.0, [12].Setpoint[40] := 30.0, [12].Setpoint[41] := 60.0, [12].Setpoint[42] := 60.0, [12].Setpoint[43] := 3000.0, [12].Setpoint[44] := 300.0, [12].Setpoint[45] := 185.0, [12].Setpoint[46] := 10.0, [12].Setpoint[47] := 25.0, [12].Setpoint[48] := 150.0, [12].Setpoint[49] := 125.0, [12].Setpoint[50] := 100.0, [12].Setpoint[51] := 80.0, [12].Setpoint[52] := 100.0, [12].Setpoint[53] := 50.0, [12].Setpoint[54] := 85.0, [12].Setpoint[55] := 40.0, [12].Setpoint[56] := 60.0, [12].Setpoint[57] := 90.0, [12].Setpoint[58] := 4.0, [12].Setpoint[61] := 10.0, [12].Setpoint[62] := 1.0, [12].Setpoint[65] := 100.0, [12].Setpoint[66] := 15.0, [12].Setpoint[67] := 50.0, [12].Setpoint[68] := 5.0, [12].Setpoint[69] := 100.0, [12].Setpoint[70] := 15.0, [12].Setpoint[71] := 100.0, [12].Setpoint[72] := 15.0, [12].Setpoint[73] := 120.0, [12].Setpoint[74] := 20.0, [12].Setpoint[75] := 120.0, [12].Setpoint[76] := 20.0, [12].Setpoint[77] := 100.0, [12].Setpoint[78] := 15.0, [12].Setpoint[79] := 100.0, [12].Setpoint[80] := 15.0, [12].Setpoint[81] := 45.0, [12].Setpoint[82] := 30.0, [12].Setpoint[83] := 5.0, [12].Setpoint[85] := 5.0, [12].Setpoint[86] := 9.0, [12].Setpoint[92] := 75.0, [12].Setpoint[93] := 90.0, [12].Setpoint[94] := 5.0, [12].Setpoint[95] := 110.0, [12].Setpoint[96] := 10.0, [12].Name := 'RECIPE #12',
        [13].Setpoint[1] := 55.0, [13].Setpoint[2] := 65.0, [13].Setpoint[3] := 60.0, [13].Setpoint[4] := 45.0, [13].Setpoint[5] := 65.0, [13].Setpoint[6] := 25.0, [13].Setpoint[7] := 53.0, [13].Setpoint[8] := 63.0, [13].Setpoint[9] := 57.0, [13].Setpoint[10] := 43.0, [13].Setpoint[11] := 63.0, [13].Setpoint[12] := 22.0, [13].Setpoint[13] := 85.0, [13].Setpoint[14] := 900.0, [13].Setpoint[15] := 300.0, [13].Setpoint[16] := 300.0, [13].Setpoint[17] := 15.0, [13].Setpoint[18] := 14.0, [13].Setpoint[19] := 15.0, [13].Setpoint[20] := 45.0, [13].Setpoint[21] := 5.0, [13].Setpoint[22] := 15.0, [13].Setpoint[23] := 300.0, [13].Setpoint[24] := 2.0, [13].Setpoint[25] := 10.0, [13].Setpoint[26] := 9.0, [13].Setpoint[27] := 10.0, [13].Setpoint[28] := 50.0, [13].Setpoint[29] := 3.0, [13].Setpoint[30] := 17.0, [13].Setpoint[31] := 300.0, [13].Setpoint[32] := 2.0, [13].Setpoint[33] := 2.0, [13].Setpoint[34] := 900.0, [13].Setpoint[37] := 70.0, [13].Setpoint[38] := 100.0, [13].Setpoint[39] := 110.0, [13].Setpoint[40] := 30.0, [13].Setpoint[41] := 60.0, [13].Setpoint[42] := 60.0, [13].Setpoint[43] := 3000.0, [13].Setpoint[44] := 300.0, [13].Setpoint[45] := 185.0, [13].Setpoint[46] := 10.0, [13].Setpoint[47] := 25.0, [13].Setpoint[48] := 150.0, [13].Setpoint[49] := 125.0, [13].Setpoint[50] := 100.0, [13].Setpoint[51] := 80.0, [13].Setpoint[52] := 100.0, [13].Setpoint[53] := 50.0, [13].Setpoint[54] := 85.0, [13].Setpoint[55] := 40.0, [13].Setpoint[56] := 60.0, [13].Setpoint[57] := 90.0, [13].Setpoint[58] := 4.0, [13].Setpoint[61] := 10.0, [13].Setpoint[62] := 1.0, [13].Setpoint[65] := 100.0, [13].Setpoint[66] := 15.0,
        [13].Setpoint[67] := 50.0, [13].Setpoint[68] := 5.0, [13].Setpoint[69] := 100.0, [13].Setpoint[70] := 15.0, [13].Setpoint[71] := 100.0, [13].Setpoint[72] := 15.0, [13].Setpoint[73] := 120.0, [13].Setpoint[74] := 20.0, [13].Setpoint[75] := 120.0, [13].Setpoint[76] := 20.0, [13].Setpoint[77] := 100.0, [13].Setpoint[78] := 15.0, [13].Setpoint[79] := 100.0, [13].Setpoint[80] := 15.0, [13].Setpoint[81] := 45.0, [13].Setpoint[82] := 30.0, [13].Setpoint[83] := 5.0, [13].Setpoint[85] := 5.0, [13].Setpoint[86] := 9.0, [13].Setpoint[92] := 75.0, [13].Setpoint[93] := 90.0, [13].Setpoint[94] := 5.0, [13].Setpoint[95] := 110.0, [13].Setpoint[96] := 10.0, [13].Name := 'RECIPE #13', [14].Setpoint[1] := 55.0, [14].Setpoint[2] := 65.0, [14].Setpoint[3] := 60.0, [14].Setpoint[4] := 45.0, [14].Setpoint[5] := 65.0, [14].Setpoint[6] := 25.0, [14].Setpoint[7] := 53.0, [14].Setpoint[8] := 63.0, [14].Setpoint[9] := 57.0, [14].Setpoint[10] := 43.0, [14].Setpoint[11] := 63.0, [14].Setpoint[12] := 22.0, [14].Setpoint[13] := 85.0, [14].Setpoint[14] := 900.0, [14].Setpoint[15] := 300.0, [14].Setpoint[16] := 300.0, [14].Setpoint[17] := 15.0, [14].Setpoint[18] := 14.0, [14].Setpoint[19] := 15.0, [14].Setpoint[20] := 45.0, [14].Setpoint[21] := 5.0, [14].Setpoint[22] := 15.0, [14].Setpoint[23] := 300.0, [14].Setpoint[24] := 2.0, [14].Setpoint[25] := 10.0, [14].Setpoint[26] := 9.0, [14].Setpoint[27] := 10.0, [14].Setpoint[28] := 50.0, [14].Setpoint[29] := 3.0, [14].Setpoint[30] := 17.0, [14].Setpoint[31] := 300.0, [14].Setpoint[32] := 2.0, [14].Setpoint[33] := 2.0, [14].Setpoint[34] := 900.0, [14].Setpoint[37] := 70.0,
        [14].Setpoint[38] := 100.0, [14].Setpoint[39] := 110.0, [14].Setpoint[40] := 30.0, [14].Setpoint[41] := 60.0, [14].Setpoint[42] := 60.0, [14].Setpoint[43] := 3000.0, [14].Setpoint[44] := 300.0, [14].Setpoint[45] := 185.0, [14].Setpoint[46] := 10.0, [14].Setpoint[47] := 25.0, [14].Setpoint[48] := 150.0, [14].Setpoint[49] := 125.0, [14].Setpoint[50] := 100.0, [14].Setpoint[51] := 80.0, [14].Setpoint[52] := 100.0, [14].Setpoint[53] := 50.0, [14].Setpoint[54] := 85.0, [14].Setpoint[55] := 40.0, [14].Setpoint[56] := 60.0, [14].Setpoint[57] := 90.0, [14].Setpoint[58] := 4.0, [14].Setpoint[61] := 10.0, [14].Setpoint[62] := 1.0, [14].Setpoint[65] := 100.0, [14].Setpoint[66] := 15.0, [14].Setpoint[67] := 50.0, [14].Setpoint[68] := 5.0, [14].Setpoint[69] := 100.0, [14].Setpoint[70] := 15.0, [14].Setpoint[71] := 100.0, [14].Setpoint[72] := 15.0, [14].Setpoint[73] := 120.0, [14].Setpoint[74] := 20.0, [14].Setpoint[75] := 120.0, [14].Setpoint[76] := 20.0, [14].Setpoint[77] := 100.0, [14].Setpoint[78] := 15.0, [14].Setpoint[79] := 100.0, [14].Setpoint[80] := 15.0, [14].Setpoint[81] := 45.0, [14].Setpoint[82] := 30.0, [14].Setpoint[83] := 5.0, [14].Setpoint[85] := 5.0, [14].Setpoint[86] := 9.0, [14].Setpoint[92] := 75.0, [14].Setpoint[93] := 90.0, [14].Setpoint[94] := 5.0, [14].Setpoint[95] := 110.0, [14].Setpoint[96] := 10.0, [14].Name := 'RECIPE #14', [15].Setpoint[1] := 55.0, [15].Setpoint[2] := 65.0, [15].Setpoint[3] := 60.0, [15].Setpoint[4] := 45.0, [15].Setpoint[5] := 65.0, [15].Setpoint[6] := 25.0, [15].Setpoint[7] := 53.0, [15].Setpoint[8] := 63.0, [15].Setpoint[9] := 57.0, [15].Setpoint[10] := 43.0,
        [15].Setpoint[11] := 63.0, [15].Setpoint[12] := 22.0, [15].Setpoint[13] := 85.0, [15].Setpoint[14] := 900.0, [15].Setpoint[15] := 300.0, [15].Setpoint[16] := 300.0, [15].Setpoint[17] := 15.0, [15].Setpoint[18] := 14.0, [15].Setpoint[19] := 15.0, [15].Setpoint[20] := 45.0, [15].Setpoint[21] := 5.0, [15].Setpoint[22] := 15.0, [15].Setpoint[23] := 300.0, [15].Setpoint[24] := 2.0, [15].Setpoint[25] := 10.0, [15].Setpoint[26] := 9.0, [15].Setpoint[27] := 10.0, [15].Setpoint[28] := 50.0, [15].Setpoint[29] := 3.0, [15].Setpoint[30] := 17.0, [15].Setpoint[31] := 300.0, [15].Setpoint[32] := 2.0, [15].Setpoint[33] := 2.0, [15].Setpoint[34] := 900.0, [15].Setpoint[37] := 70.0, [15].Setpoint[38] := 100.0, [15].Setpoint[39] := 110.0, [15].Setpoint[40] := 30.0, [15].Setpoint[41] := 60.0, [15].Setpoint[42] := 60.0, [15].Setpoint[43] := 3000.0, [15].Setpoint[44] := 300.0, [15].Setpoint[45] := 185.0, [15].Setpoint[46] := 10.0, [15].Setpoint[47] := 25.0, [15].Setpoint[48] := 150.0, [15].Setpoint[49] := 125.0, [15].Setpoint[50] := 100.0, [15].Setpoint[51] := 80.0, [15].Setpoint[52] := 100.0, [15].Setpoint[53] := 50.0, [15].Setpoint[54] := 85.0, [15].Setpoint[55] := 40.0, [15].Setpoint[56] := 60.0, [15].Setpoint[57] := 90.0, [15].Setpoint[58] := 4.0, [15].Setpoint[61] := 10.0, [15].Setpoint[62] := 1.0, [15].Setpoint[65] := 100.0, [15].Setpoint[66] := 15.0, [15].Setpoint[67] := 50.0, [15].Setpoint[68] := 5.0, [15].Setpoint[69] := 100.0, [15].Setpoint[70] := 15.0, [15].Setpoint[71] := 100.0, [15].Setpoint[72] := 15.0, [15].Setpoint[73] := 120.0, [15].Setpoint[74] := 20.0, [15].Setpoint[75] := 120.0, [15].Setpoint[76] := 20.0,
        [15].Setpoint[77] := 100.0, [15].Setpoint[78] := 15.0, [15].Setpoint[79] := 100.0, [15].Setpoint[80] := 15.0, [15].Setpoint[81] := 45.0, [15].Setpoint[82] := 30.0, [15].Setpoint[83] := 5.0, [15].Setpoint[85] := 5.0, [15].Setpoint[86] := 9.0, [15].Setpoint[92] := 75.0, [15].Setpoint[93] := 90.0, [15].Setpoint[94] := 5.0, [15].Setpoint[95] := 110.0, [15].Setpoint[96] := 10.0, [15].Name := 'RECIPE #15', [16].Setpoint[1] := 55.0, [16].Setpoint[2] := 65.0, [16].Setpoint[3] := 60.0, [16].Setpoint[4] := 45.0, [16].Setpoint[5] := 65.0, [16].Setpoint[6] := 25.0, [16].Setpoint[7] := 53.0, [16].Setpoint[8] := 63.0, [16].Setpoint[9] := 57.0, [16].Setpoint[10] := 43.0, [16].Setpoint[11] := 63.0, [16].Setpoint[12] := 22.0, [16].Setpoint[13] := 85.0, [16].Setpoint[14] := 900.0, [16].Setpoint[15] := 300.0, [16].Setpoint[16] := 300.0, [16].Setpoint[17] := 15.0, [16].Setpoint[18] := 14.0, [16].Setpoint[19] := 15.0, [16].Setpoint[20] := 45.0, [16].Setpoint[21] := 5.0, [16].Setpoint[22] := 15.0, [16].Setpoint[23] := 300.0, [16].Setpoint[24] := 2.0, [16].Setpoint[25] := 10.0, [16].Setpoint[26] := 9.0, [16].Setpoint[27] := 10.0, [16].Setpoint[28] := 50.0, [16].Setpoint[29] := 3.0, [16].Setpoint[30] := 17.0, [16].Setpoint[31] := 300.0, [16].Setpoint[32] := 2.0, [16].Setpoint[33] := 2.0, [16].Setpoint[34] := 900.0, [16].Setpoint[37] := 70.0, [16].Setpoint[38] := 100.0, [16].Setpoint[39] := 110.0, [16].Setpoint[40] := 30.0, [16].Setpoint[41] := 60.0, [16].Setpoint[42] := 60.0, [16].Setpoint[43] := 3000.0, [16].Setpoint[44] := 300.0, [16].Setpoint[45] := 185.0, [16].Setpoint[46] := 10.0, [16].Setpoint[47] := 25.0,
        [16].Setpoint[48] := 150.0, [16].Setpoint[49] := 125.0, [16].Setpoint[50] := 100.0, [16].Setpoint[51] := 80.0, [16].Setpoint[52] := 100.0, [16].Setpoint[53] := 50.0, [16].Setpoint[54] := 85.0, [16].Setpoint[55] := 40.0, [16].Setpoint[56] := 60.0, [16].Setpoint[57] := 90.0, [16].Setpoint[58] := 4.0, [16].Setpoint[61] := 10.0, [16].Setpoint[62] := 1.0, [16].Setpoint[65] := 100.0, [16].Setpoint[66] := 15.0, [16].Setpoint[67] := 50.0, [16].Setpoint[68] := 5.0, [16].Setpoint[69] := 100.0, [16].Setpoint[70] := 15.0, [16].Setpoint[71] := 100.0, [16].Setpoint[72] := 15.0, [16].Setpoint[73] := 120.0, [16].Setpoint[74] := 20.0, [16].Setpoint[75] := 120.0, [16].Setpoint[76] := 20.0, [16].Setpoint[77] := 100.0, [16].Setpoint[78] := 15.0, [16].Setpoint[79] := 100.0, [16].Setpoint[80] := 15.0, [16].Setpoint[81] := 45.0, [16].Setpoint[82] := 30.0, [16].Setpoint[83] := 5.0, [16].Setpoint[85] := 5.0, [16].Setpoint[86] := 9.0, [16].Setpoint[92] := 75.0, [16].Setpoint[93] := 90.0, [16].Setpoint[94] := 5.0, [16].Setpoint[95] := 110.0, [16].Setpoint[96] := 10.0, [16].Name := 'RECIPE #16', [17].Setpoint[1] := 55.0, [17].Setpoint[2] := 65.0, [17].Setpoint[3] := 60.0, [17].Setpoint[4] := 45.0, [17].Setpoint[5] := 65.0, [17].Setpoint[6] := 25.0, [17].Setpoint[7] := 53.0, [17].Setpoint[8] := 63.0, [17].Setpoint[9] := 57.0, [17].Setpoint[10] := 43.0, [17].Setpoint[11] := 63.0, [17].Setpoint[12] := 22.0, [17].Setpoint[13] := 85.0, [17].Setpoint[14] := 900.0, [17].Setpoint[15] := 300.0, [17].Setpoint[16] := 300.0, [17].Setpoint[17] := 15.0, [17].Setpoint[18] := 14.0, [17].Setpoint[19] := 15.0, [17].Setpoint[20] := 45.0,
        [17].Setpoint[21] := 5.0, [17].Setpoint[22] := 15.0, [17].Setpoint[23] := 300.0, [17].Setpoint[24] := 2.0, [17].Setpoint[25] := 10.0, [17].Setpoint[26] := 9.0, [17].Setpoint[27] := 10.0, [17].Setpoint[28] := 50.0, [17].Setpoint[29] := 3.0, [17].Setpoint[30] := 17.0, [17].Setpoint[31] := 300.0, [17].Setpoint[32] := 2.0, [17].Setpoint[33] := 2.0, [17].Setpoint[34] := 900.0, [17].Setpoint[37] := 70.0, [17].Setpoint[38] := 100.0, [17].Setpoint[39] := 110.0, [17].Setpoint[40] := 30.0, [17].Setpoint[41] := 60.0, [17].Setpoint[42] := 60.0, [17].Setpoint[43] := 3000.0, [17].Setpoint[44] := 300.0, [17].Setpoint[45] := 185.0, [17].Setpoint[46] := 10.0, [17].Setpoint[47] := 25.0, [17].Setpoint[48] := 150.0, [17].Setpoint[49] := 125.0, [17].Setpoint[50] := 100.0, [17].Setpoint[51] := 80.0, [17].Setpoint[52] := 100.0, [17].Setpoint[53] := 50.0, [17].Setpoint[54] := 85.0, [17].Setpoint[55] := 40.0, [17].Setpoint[56] := 60.0, [17].Setpoint[57] := 90.0, [17].Setpoint[58] := 4.0, [17].Setpoint[61] := 10.0, [17].Setpoint[62] := 1.0, [17].Setpoint[65] := 100.0, [17].Setpoint[66] := 15.0, [17].Setpoint[67] := 50.0, [17].Setpoint[68] := 5.0, [17].Setpoint[69] := 100.0, [17].Setpoint[70] := 15.0, [17].Setpoint[71] := 100.0, [17].Setpoint[72] := 15.0, [17].Setpoint[73] := 120.0, [17].Setpoint[74] := 20.0, [17].Setpoint[75] := 120.0, [17].Setpoint[76] := 20.0, [17].Setpoint[77] := 100.0, [17].Setpoint[78] := 15.0, [17].Setpoint[79] := 100.0, [17].Setpoint[80] := 15.0, [17].Setpoint[81] := 45.0, [17].Setpoint[82] := 30.0, [17].Setpoint[83] := 5.0, [17].Setpoint[85] := 5.0, [17].Setpoint[86] := 9.0, [17].Setpoint[92] := 75.0,
        [17].Setpoint[93] := 90.0, [17].Setpoint[94] := 5.0, [17].Setpoint[95] := 110.0, [17].Setpoint[96] := 10.0, [17].Name := 'RECIPE #17', [18].Setpoint[1] := 55.0, [18].Setpoint[2] := 65.0, [18].Setpoint[3] := 60.0, [18].Setpoint[4] := 45.0, [18].Setpoint[5] := 65.0, [18].Setpoint[6] := 25.0, [18].Setpoint[7] := 53.0, [18].Setpoint[8] := 63.0, [18].Setpoint[9] := 57.0, [18].Setpoint[10] := 43.0, [18].Setpoint[11] := 63.0, [18].Setpoint[12] := 22.0, [18].Setpoint[13] := 85.0, [18].Setpoint[14] := 900.0, [18].Setpoint[15] := 300.0, [18].Setpoint[16] := 300.0, [18].Setpoint[17] := 15.0, [18].Setpoint[18] := 14.0, [18].Setpoint[19] := 15.0, [18].Setpoint[20] := 45.0, [18].Setpoint[21] := 5.0, [18].Setpoint[22] := 15.0, [18].Setpoint[23] := 300.0, [18].Setpoint[24] := 2.0, [18].Setpoint[25] := 10.0, [18].Setpoint[26] := 9.0, [18].Setpoint[27] := 10.0, [18].Setpoint[28] := 50.0, [18].Setpoint[29] := 3.0, [18].Setpoint[30] := 17.0, [18].Setpoint[31] := 300.0, [18].Setpoint[32] := 2.0, [18].Setpoint[33] := 2.0, [18].Setpoint[34] := 900.0, [18].Setpoint[37] := 70.0, [18].Setpoint[38] := 100.0, [18].Setpoint[39] := 110.0, [18].Setpoint[40] := 30.0, [18].Setpoint[41] := 60.0, [18].Setpoint[42] := 60.0, [18].Setpoint[43] := 3000.0, [18].Setpoint[44] := 300.0, [18].Setpoint[45] := 185.0, [18].Setpoint[46] := 10.0, [18].Setpoint[47] := 25.0, [18].Setpoint[48] := 150.0, [18].Setpoint[49] := 125.0, [18].Setpoint[50] := 100.0, [18].Setpoint[51] := 80.0, [18].Setpoint[52] := 100.0, [18].Setpoint[53] := 50.0, [18].Setpoint[54] := 85.0, [18].Setpoint[55] := 40.0, [18].Setpoint[56] := 60.0, [18].Setpoint[57] := 90.0,
        [18].Setpoint[58] := 4.0, [18].Setpoint[61] := 10.0, [18].Setpoint[62] := 1.0, [18].Setpoint[65] := 100.0, [18].Setpoint[66] := 15.0, [18].Setpoint[67] := 50.0, [18].Setpoint[68] := 5.0, [18].Setpoint[69] := 100.0, [18].Setpoint[70] := 15.0, [18].Setpoint[71] := 100.0, [18].Setpoint[72] := 15.0, [18].Setpoint[73] := 120.0, [18].Setpoint[74] := 20.0, [18].Setpoint[75] := 120.0, [18].Setpoint[76] := 20.0, [18].Setpoint[77] := 100.0, [18].Setpoint[78] := 15.0, [18].Setpoint[79] := 100.0, [18].Setpoint[80] := 15.0, [18].Setpoint[81] := 45.0, [18].Setpoint[82] := 30.0, [18].Setpoint[83] := 5.0, [18].Setpoint[85] := 5.0, [18].Setpoint[86] := 9.0, [18].Setpoint[92] := 75.0, [18].Setpoint[93] := 90.0, [18].Setpoint[94] := 5.0, [18].Setpoint[95] := 110.0, [18].Setpoint[96] := 10.0, [18].Name := 'RECIPE #18', [19].Setpoint[1] := 55.0, [19].Setpoint[2] := 65.0, [19].Setpoint[3] := 60.0, [19].Setpoint[4] := 45.0, [19].Setpoint[5] := 65.0, [19].Setpoint[6] := 25.0, [19].Setpoint[7] := 53.0, [19].Setpoint[8] := 63.0, [19].Setpoint[9] := 57.0, [19].Setpoint[10] := 43.0, [19].Setpoint[11] := 63.0, [19].Setpoint[12] := 22.0, [19].Setpoint[13] := 85.0, [19].Setpoint[14] := 900.0, [19].Setpoint[15] := 300.0, [19].Setpoint[16] := 300.0, [19].Setpoint[17] := 15.0, [19].Setpoint[18] := 14.0, [19].Setpoint[19] := 15.0, [19].Setpoint[20] := 45.0, [19].Setpoint[21] := 5.0, [19].Setpoint[22] := 15.0, [19].Setpoint[23] := 300.0, [19].Setpoint[24] := 2.0, [19].Setpoint[25] := 10.0, [19].Setpoint[26] := 9.0, [19].Setpoint[27] := 10.0, [19].Setpoint[28] := 50.0, [19].Setpoint[29] := 3.0, [19].Setpoint[30] := 17.0,
        [19].Setpoint[31] := 300.0, [19].Setpoint[32] := 2.0, [19].Setpoint[33] := 2.0, [19].Setpoint[34] := 900.0, [19].Setpoint[37] := 70.0, [19].Setpoint[38] := 100.0, [19].Setpoint[39] := 110.0, [19].Setpoint[40] := 30.0, [19].Setpoint[41] := 60.0, [19].Setpoint[42] := 60.0, [19].Setpoint[43] := 3000.0, [19].Setpoint[44] := 300.0, [19].Setpoint[45] := 185.0, [19].Setpoint[46] := 10.0, [19].Setpoint[47] := 25.0, [19].Setpoint[48] := 150.0, [19].Setpoint[49] := 125.0, [19].Setpoint[50] := 100.0, [19].Setpoint[51] := 80.0, [19].Setpoint[52] := 100.0, [19].Setpoint[53] := 50.0, [19].Setpoint[54] := 85.0, [19].Setpoint[55] := 40.0, [19].Setpoint[56] := 60.0, [19].Setpoint[57] := 90.0, [19].Setpoint[58] := 4.0, [19].Setpoint[61] := 10.0, [19].Setpoint[62] := 1.0, [19].Setpoint[65] := 100.0, [19].Setpoint[66] := 15.0, [19].Setpoint[67] := 50.0, [19].Setpoint[68] := 5.0, [19].Setpoint[69] := 100.0, [19].Setpoint[70] := 15.0, [19].Setpoint[71] := 100.0, [19].Setpoint[72] := 15.0, [19].Setpoint[73] := 120.0, [19].Setpoint[74] := 20.0, [19].Setpoint[75] := 120.0, [19].Setpoint[76] := 20.0, [19].Setpoint[77] := 100.0, [19].Setpoint[78] := 15.0, [19].Setpoint[79] := 100.0, [19].Setpoint[80] := 15.0, [19].Setpoint[81] := 45.0, [19].Setpoint[82] := 30.0, [19].Setpoint[83] := 5.0, [19].Setpoint[85] := 5.0, [19].Setpoint[86] := 9.0, [19].Setpoint[92] := 75.0, [19].Setpoint[93] := 90.0, [19].Setpoint[94] := 5.0, [19].Setpoint[95] := 110.0, [19].Setpoint[96] := 10.0, [19].Name := 'RECIPE #19', [20].Setpoint[1] := 55.0, [20].Setpoint[2] := 65.0, [20].Setpoint[3] := 60.0, [20].Setpoint[4] := 45.0, [20].Setpoint[5] := 65.0,
        [20].Setpoint[6] := 25.0, [20].Setpoint[7] := 53.0, [20].Setpoint[8] := 63.0, [20].Setpoint[9] := 57.0, [20].Setpoint[10] := 43.0, [20].Setpoint[11] := 63.0, [20].Setpoint[12] := 22.0, [20].Setpoint[13] := 85.0, [20].Setpoint[14] := 900.0, [20].Setpoint[15] := 300.0, [20].Setpoint[16] := 300.0, [20].Setpoint[17] := 15.0, [20].Setpoint[18] := 14.0, [20].Setpoint[19] := 15.0, [20].Setpoint[20] := 45.0, [20].Setpoint[21] := 5.0, [20].Setpoint[22] := 15.0, [20].Setpoint[23] := 300.0, [20].Setpoint[24] := 2.0, [20].Setpoint[25] := 10.0, [20].Setpoint[26] := 9.0, [20].Setpoint[27] := 10.0, [20].Setpoint[28] := 50.0, [20].Setpoint[29] := 3.0, [20].Setpoint[30] := 17.0, [20].Setpoint[31] := 300.0, [20].Setpoint[32] := 2.0, [20].Setpoint[33] := 2.0, [20].Setpoint[34] := 900.0, [20].Setpoint[37] := 70.0, [20].Setpoint[38] := 100.0, [20].Setpoint[39] := 110.0, [20].Setpoint[40] := 30.0, [20].Setpoint[41] := 60.0, [20].Setpoint[42] := 60.0, [20].Setpoint[43] := 3000.0, [20].Setpoint[44] := 300.0, [20].Setpoint[45] := 185.0, [20].Setpoint[46] := 10.0, [20].Setpoint[47] := 25.0, [20].Setpoint[48] := 150.0, [20].Setpoint[49] := 125.0, [20].Setpoint[50] := 100.0, [20].Setpoint[51] := 80.0, [20].Setpoint[52] := 100.0, [20].Setpoint[53] := 50.0, [20].Setpoint[54] := 85.0, [20].Setpoint[55] := 40.0, [20].Setpoint[56] := 60.0, [20].Setpoint[57] := 90.0, [20].Setpoint[58] := 4.0, [20].Setpoint[61] := 10.0, [20].Setpoint[62] := 1.0, [20].Setpoint[65] := 100.0, [20].Setpoint[66] := 15.0, [20].Setpoint[67] := 50.0, [20].Setpoint[68] := 5.0, [20].Setpoint[69] := 100.0, [20].Setpoint[70] := 15.0, [20].Setpoint[71] := 100.0,
        [20].Setpoint[72] := 15.0, [20].Setpoint[73] := 120.0, [20].Setpoint[74] := 20.0, [20].Setpoint[75] := 120.0, [20].Setpoint[76] := 20.0, [20].Setpoint[77] := 100.0, [20].Setpoint[78] := 15.0, [20].Setpoint[79] := 100.0, [20].Setpoint[80] := 15.0, [20].Setpoint[81] := 45.0, [20].Setpoint[82] := 30.0, [20].Setpoint[83] := 5.0, [20].Setpoint[85] := 5.0, [20].Setpoint[86] := 9.0, [20].Setpoint[92] := 75.0, [20].Setpoint[93] := 90.0, [20].Setpoint[94] := 5.0, [20].Setpoint[95] := 110.0, [20].Setpoint[96] := 10.0, [20].Name := 'RECIPE #20', [21].Setpoint[1] := 55.0, [21].Setpoint[2] := 65.0, [21].Setpoint[3] := 60.0, [21].Setpoint[4] := 45.0, [21].Setpoint[5] := 65.0, [21].Setpoint[6] := 25.0, [21].Setpoint[7] := 53.0, [21].Setpoint[8] := 63.0, [21].Setpoint[9] := 57.0, [21].Setpoint[10] := 43.0, [21].Setpoint[11] := 63.0, [21].Setpoint[12] := 22.0, [21].Setpoint[13] := 85.0, [21].Setpoint[14] := 900.0, [21].Setpoint[15] := 300.0, [21].Setpoint[16] := 300.0, [21].Setpoint[17] := 15.0, [21].Setpoint[18] := 14.0, [21].Setpoint[19] := 15.0, [21].Setpoint[20] := 45.0, [21].Setpoint[21] := 5.0, [21].Setpoint[22] := 15.0, [21].Setpoint[23] := 300.0, [21].Setpoint[24] := 2.0, [21].Setpoint[25] := 10.0, [21].Setpoint[26] := 9.0, [21].Setpoint[27] := 10.0, [21].Setpoint[28] := 50.0, [21].Setpoint[29] := 3.0, [21].Setpoint[30] := 17.0, [21].Setpoint[31] := 300.0, [21].Setpoint[32] := 2.0, [21].Setpoint[33] := 2.0, [21].Setpoint[34] := 900.0, [21].Setpoint[37] := 70.0, [21].Setpoint[38] := 100.0, [21].Setpoint[39] := 110.0, [21].Setpoint[40] := 30.0, [21].Setpoint[41] := 60.0, [21].Setpoint[42] := 60.0,
        [21].Setpoint[43] := 3000.0, [21].Setpoint[44] := 300.0, [21].Setpoint[45] := 185.0, [21].Setpoint[46] := 10.0, [21].Setpoint[47] := 25.0, [21].Setpoint[48] := 150.0, [21].Setpoint[49] := 125.0, [21].Setpoint[50] := 100.0, [21].Setpoint[51] := 80.0, [21].Setpoint[52] := 100.0, [21].Setpoint[53] := 50.0, [21].Setpoint[54] := 85.0, [21].Setpoint[55] := 40.0, [21].Setpoint[56] := 60.0, [21].Setpoint[57] := 90.0, [21].Setpoint[58] := 4.0, [21].Setpoint[61] := 10.0, [21].Setpoint[62] := 1.0, [21].Setpoint[65] := 100.0, [21].Setpoint[66] := 15.0, [21].Setpoint[67] := 50.0, [21].Setpoint[68] := 5.0, [21].Setpoint[69] := 100.0, [21].Setpoint[70] := 15.0, [21].Setpoint[71] := 100.0, [21].Setpoint[72] := 15.0, [21].Setpoint[73] := 120.0, [21].Setpoint[74] := 20.0, [21].Setpoint[75] := 120.0, [21].Setpoint[76] := 20.0, [21].Setpoint[77] := 100.0, [21].Setpoint[78] := 15.0, [21].Setpoint[79] := 100.0, [21].Setpoint[80] := 15.0, [21].Setpoint[81] := 45.0, [21].Setpoint[82] := 30.0, [21].Setpoint[83] := 5.0, [21].Setpoint[85] := 5.0, [21].Setpoint[86] := 9.0, [21].Setpoint[92] := 75.0, [21].Setpoint[93] := 90.0, [21].Setpoint[94] := 5.0, [21].Setpoint[95] := 110.0, [21].Setpoint[96] := 10.0, [21].Name := 'RECIPE #21', [22].Setpoint[1] := 55.0, [22].Setpoint[2] := 65.0, [22].Setpoint[3] := 60.0, [22].Setpoint[4] := 45.0, [22].Setpoint[5] := 65.0, [22].Setpoint[6] := 25.0, [22].Setpoint[7] := 53.0, [22].Setpoint[8] := 63.0, [22].Setpoint[9] := 57.0, [22].Setpoint[10] := 43.0, [22].Setpoint[11] := 63.0, [22].Setpoint[12] := 22.0, [22].Setpoint[13] := 85.0, [22].Setpoint[14] := 900.0, [22].Setpoint[15] := 300.0,
        [22].Setpoint[16] := 300.0, [22].Setpoint[17] := 15.0, [22].Setpoint[18] := 14.0, [22].Setpoint[19] := 15.0, [22].Setpoint[20] := 45.0, [22].Setpoint[21] := 5.0, [22].Setpoint[22] := 15.0, [22].Setpoint[23] := 300.0, [22].Setpoint[24] := 2.0, [22].Setpoint[25] := 10.0, [22].Setpoint[26] := 9.0, [22].Setpoint[27] := 10.0, [22].Setpoint[28] := 50.0, [22].Setpoint[29] := 3.0, [22].Setpoint[30] := 17.0, [22].Setpoint[31] := 300.0, [22].Setpoint[32] := 2.0, [22].Setpoint[33] := 2.0, [22].Setpoint[34] := 900.0, [22].Setpoint[37] := 70.0, [22].Setpoint[38] := 100.0, [22].Setpoint[39] := 110.0, [22].Setpoint[40] := 30.0, [22].Setpoint[41] := 60.0, [22].Setpoint[42] := 60.0, [22].Setpoint[43] := 3000.0, [22].Setpoint[44] := 300.0, [22].Setpoint[45] := 185.0, [22].Setpoint[46] := 10.0, [22].Setpoint[47] := 25.0, [22].Setpoint[48] := 150.0, [22].Setpoint[49] := 125.0, [22].Setpoint[50] := 100.0, [22].Setpoint[51] := 80.0, [22].Setpoint[52] := 100.0, [22].Setpoint[53] := 50.0, [22].Setpoint[54] := 85.0, [22].Setpoint[55] := 40.0, [22].Setpoint[56] := 60.0, [22].Setpoint[57] := 90.0, [22].Setpoint[58] := 4.0, [22].Setpoint[61] := 10.0, [22].Setpoint[62] := 1.0, [22].Setpoint[65] := 100.0, [22].Setpoint[66] := 15.0, [22].Setpoint[67] := 50.0, [22].Setpoint[68] := 5.0, [22].Setpoint[69] := 100.0, [22].Setpoint[70] := 15.0, [22].Setpoint[71] := 100.0, [22].Setpoint[72] := 15.0, [22].Setpoint[73] := 120.0, [22].Setpoint[74] := 20.0, [22].Setpoint[75] := 120.0, [22].Setpoint[76] := 20.0, [22].Setpoint[77] := 100.0, [22].Setpoint[78] := 15.0, [22].Setpoint[79] := 100.0, [22].Setpoint[80] := 15.0, [22].Setpoint[81] := 45.0,
        [22].Setpoint[82] := 30.0, [22].Setpoint[83] := 5.0, [22].Setpoint[85] := 5.0, [22].Setpoint[86] := 9.0, [22].Setpoint[92] := 75.0, [22].Setpoint[93] := 90.0, [22].Setpoint[94] := 5.0, [22].Setpoint[95] := 110.0, [22].Setpoint[96] := 10.0, [22].Name := 'RECIPE #22', [23].Setpoint[1] := 55.0, [23].Setpoint[2] := 65.0, [23].Setpoint[3] := 60.0, [23].Setpoint[4] := 45.0, [23].Setpoint[5] := 65.0, [23].Setpoint[6] := 25.0, [23].Setpoint[7] := 53.0, [23].Setpoint[8] := 63.0, [23].Setpoint[9] := 57.0, [23].Setpoint[10] := 43.0, [23].Setpoint[11] := 63.0, [23].Setpoint[12] := 22.0, [23].Setpoint[13] := 85.0, [23].Setpoint[14] := 900.0, [23].Setpoint[15] := 300.0, [23].Setpoint[16] := 300.0, [23].Setpoint[17] := 15.0, [23].Setpoint[18] := 14.0, [23].Setpoint[19] := 15.0, [23].Setpoint[20] := 45.0, [23].Setpoint[21] := 5.0, [23].Setpoint[22] := 15.0, [23].Setpoint[23] := 300.0, [23].Setpoint[24] := 2.0, [23].Setpoint[25] := 10.0, [23].Setpoint[26] := 9.0, [23].Setpoint[27] := 10.0, [23].Setpoint[28] := 50.0, [23].Setpoint[29] := 3.0, [23].Setpoint[30] := 17.0, [23].Setpoint[31] := 300.0, [23].Setpoint[32] := 2.0, [23].Setpoint[33] := 2.0, [23].Setpoint[34] := 900.0, [23].Setpoint[37] := 70.0, [23].Setpoint[38] := 100.0, [23].Setpoint[39] := 110.0, [23].Setpoint[40] := 30.0, [23].Setpoint[41] := 60.0, [23].Setpoint[42] := 60.0, [23].Setpoint[43] := 3000.0, [23].Setpoint[44] := 300.0, [23].Setpoint[45] := 185.0, [23].Setpoint[46] := 10.0, [23].Setpoint[47] := 25.0, [23].Setpoint[48] := 150.0, [23].Setpoint[49] := 125.0, [23].Setpoint[50] := 100.0, [23].Setpoint[51] := 80.0, [23].Setpoint[52] := 100.0,
        [23].Setpoint[53] := 50.0, [23].Setpoint[54] := 85.0, [23].Setpoint[55] := 40.0, [23].Setpoint[56] := 60.0, [23].Setpoint[57] := 90.0, [23].Setpoint[58] := 4.0, [23].Setpoint[61] := 10.0, [23].Setpoint[62] := 1.0, [23].Setpoint[65] := 100.0, [23].Setpoint[66] := 15.0, [23].Setpoint[67] := 50.0, [23].Setpoint[68] := 5.0, [23].Setpoint[69] := 100.0, [23].Setpoint[70] := 15.0, [23].Setpoint[71] := 100.0, [23].Setpoint[72] := 15.0, [23].Setpoint[73] := 120.0, [23].Setpoint[74] := 20.0, [23].Setpoint[75] := 120.0, [23].Setpoint[76] := 20.0, [23].Setpoint[77] := 100.0, [23].Setpoint[78] := 15.0, [23].Setpoint[79] := 100.0, [23].Setpoint[80] := 15.0, [23].Setpoint[81] := 45.0, [23].Setpoint[82] := 30.0, [23].Setpoint[83] := 5.0, [23].Setpoint[85] := 5.0, [23].Setpoint[86] := 9.0, [23].Setpoint[92] := 75.0, [23].Setpoint[93] := 90.0, [23].Setpoint[94] := 5.0, [23].Setpoint[95] := 110.0, [23].Setpoint[96] := 10.0, [23].Name := 'RECIPE #23', [24].Setpoint[1] := 55.0, [24].Setpoint[2] := 65.0, [24].Setpoint[3] := 60.0, [24].Setpoint[4] := 45.0, [24].Setpoint[5] := 65.0, [24].Setpoint[6] := 25.0, [24].Setpoint[7] := 53.0, [24].Setpoint[8] := 63.0, [24].Setpoint[9] := 57.0, [24].Setpoint[10] := 43.0, [24].Setpoint[11] := 63.0, [24].Setpoint[12] := 22.0, [24].Setpoint[13] := 85.0, [24].Setpoint[14] := 900.0, [24].Setpoint[15] := 300.0, [24].Setpoint[16] := 300.0, [24].Setpoint[17] := 15.0, [24].Setpoint[18] := 14.0, [24].Setpoint[19] := 15.0, [24].Setpoint[20] := 45.0, [24].Setpoint[21] := 5.0, [24].Setpoint[22] := 15.0, [24].Setpoint[23] := 300.0, [24].Setpoint[24] := 2.0, [24].Setpoint[25] := 10.0,
